Gr05Auto(bEnable := TRUE);			(* Call Program *)
Gr05Home(bEnable := TRUE);			(* Call Program *)
Gr05Manual(bEnable := TRUE);			(* Call Program *)

END_PROGRAM

// ---- POUs/Machine/Group_0500 - Transport/Gr05MachineMode/Gr05Auto/Gr05Auto.TcPOU
PROGRAM Gr05Auto
VAR_INPUT
	(* Input variables / Eingang Variablen *)
	bEnable					:BOOL;						(* Enable Gr05Auto *)
	bExecute				:BOOL;						(* Auto execute *)

	(* Instances *)
	fbInit						:FB_Gr05AutoInit;
	fbProcedure				:FB_Gr05AutoProcedure;

END_VAR
VAR
	(* Enummerations *)

	(* Variables *)
	SFCCurrentStepHis			:ARRAY[0..120] OF STRING;
	bClearHis						:BOOL;
	usnt : INT := 1;
	(* References *)

	(* Interfaces *)

	(* Instances *)
	rtExecute					:R_TRIG;
	fbAlarm					:FB_Gr05AutoAlarm;
END_VAR
VAR CONSTANT
	nFatalErrorMaxIdx				:INT := 0;						(* Maximal index of  using alarms *)
	nErrorMaxIdx					:INT := 2;						(* Maximal index of  using alarms *)
	nWarningMaxIdx				:INT := 1;						(* Maximal index of  using alarms *)
	nMessageMaxIdx				:INT := 0;						(* Maximal index of  using alarms *)
	nHintMaxIdx					:INT := 0;						(* Maximal index of  using alarms *)

	dnFatalErrorBaseIdentNo		:DINT := 52000;				(* Fatal error identification number *)
	dnErrorBaseIdentNo			:DINT := 52100;				(* Error identification number *)
	dnWarningBaseIdentNo		:DINT := 52200;				(* Warning identification number *)
	dnMessageBaseIdentNo		:DINT := 52300;				(* Message identification number *)
	dnHintBaseIdentNo			:DINT := 52400;				(* Hint identification number *)
END_VAR

IF NOT bEnable
THEN
    RETURN;
END_IF;

(* Check auto execute *)
bExecute := bgGr00ModeAutomatic
		     AND NOT fbInit.bFirstTime;

rtExecute(CLK := bExecute);

IF rtExecute.Q
THEN
	A_Init();
END_IF;

A_Procedure();
A_Functions();
A_Alarm();

ACTION A_Alarm:

(* Collect and execute input alarms *)
fbAlarm.stAlarmIn.arbError[0].bActive := fbProcedure.bErrorPipeBeginNoDetected;
fbAlarm.stAlarmIn.arbError[0].dnCode := dnErrorBaseIdentNo + 0;

fbAlarm.stAlarmIn.arbError[1].bActive := fbProcedure.bErrorPipeEndNoDetected;
fbAlarm.stAlarmIn.arbError[1].dnCode := dnErrorBaseIdentNo + 1;

fbAlarm.stAlarmIn.arbError[2].bActive := fbProcedure.bErrorCollisionDetected;
fbAlarm.stAlarmIn.arbError[2].dnCode := dnErrorBaseIdentNo + 2;

fbAlarm.stAlarmIn.arbWarning[0].bActive := fbProcedure.bWarningPipeBeginNoDetected;
fbAlarm.stAlarmIn.arbWarning[0].dnCode := dnWarningBaseIdentNo + 0;

fbAlarm(
	etMachineMode := etgGr00MachineMode,
	etMachineState := etgGr00MachineState,
	bNoEStop := bgGr00NoEmergencyStop,
	bConfirmAlarm := bgGr00ConfirmAlarm,
	dtDateTime := stgGr00DateTime.dtDateTime,
	nFatalErrorMaxIdx := nFatalErrorMaxIdx,
	nErrorMaxIdx := nErrorMaxIdx,
	nWarningMaxIdx := nWarningMaxIdx,
	nMessageMaxIdx := nMessageMaxIdx,
	nHintMaxIdx := nHintMaxIdx,
	bMoveInterrupted := bgGr05MoveInterrupted,
	bHomeCompleted := bgGr05HomeCompleted,
	stAlarmOut => stgGr05Alarm.stAuto
);
END_ACTION

ACTION A_Functions:

;
END_ACTION

ACTION A_Init:

(* Initializing variables *)
fbInit();
END_ACTION

ACTION A_Procedure:

(* Execute auto procedure *)
fbProcedure(
	bEnable := fbInit.bFirstTime,
	bExecute := bgGr05StartProcess,
	bInterrupt := FALSE(*NOT bgGr05StartProcess*),
	bReleaseNextStep := bgGr05StartProcess,
	bDone => bgGr05AutoCompleted,
	bInterrupted => bgGr05MoveInterrupted
);



(* This loup used to track the steps of this sequence *)
IF bClearHis THEN
	FOR usnt := 120 TO 1 BY  -1  DO
		SFCCurrentStepHis[usnt] := '' ;
	END_FOR
	bClearHis := FALSE;
ELSIF  fbProcedure.SFCCurrentStep <> SFCCurrentStepHis[0]  THEN
	FOR usnt := 120 TO 1 BY  -1  DO
		SFCCurrentStepHis[usnt] := SFCCurrentStepHis[usnt - 1] ;
	END_FOR
		SFCCurrentStepHis[0] := fbProcedure.SFCCurrentStep;
END_IF
END_ACTION

END_PROGRAM

// ---- POUs/Machine/Group_0500 - Transport/Gr05MachineMode/Gr05Home/Gr05Home.TcPOU
PROGRAM Gr05Home
VAR_INPUT
	(* Input variables / Eingang Variablen *)
	bEnable					:BOOL;						(* Enable Gr02Home *)
	bExecute				:BOOL;						(* Home execute *)

	(* Instances *)
	fbInit						:FB_Gr05HomeInit;
	fbProcedure				:FB_Gr05HomeProcedure;

	fbAxisClamp1				:FB_Gr05HomeAxisClamp1;
	fbAxisClamp2				:FB_Gr05HomeAxisClamp2;

END_VAR
VAR
	(* Enummerations *)

	(* Variables *)

	(* References *)

	(* Interfaces *)

	(* Instances *)
	rtExecute					:R_TRIG;

	fbAlarm					:FB_Gr05HomeAlarm;

END_VAR
VAR CONSTANT
	nFatalErrorMaxIdx				:INT := 0;						(* Maximal index of  using alarms *)
	nErrorMaxIdx					:INT := 2;						(* Maximal index of  using alarms *)
	nWarningMaxIdx				:INT := 0;						(* Maximal index of  using alarms *)
	nMessageMaxIdx				:INT := 0;						(* Maximal index of  using alarms *)
	nHintMaxIdx					:INT := 0;						(* Maximal index of  using alarms *)

	dnFatalErrorBaseIdentNo		:DINT := 53000;					(* Fatal error identification number *)
	dnErrorBaseIdentNo			:DINT := 53100;					(* Error identification number *)	
	dnWarningBaseIdentNo		:DINT := 53200;					(* Warning identification number *)	
	dnMessageBaseIdentNo		:DINT := 53300;					(* Message identification number *)	
	dnHintBaseIdentNo			:DINT := 53400;					(* Hint identification number *)
END_VAR

IF NOT bEnable
THEN
	RETURN;
END_IF;

(* Check home execute *)
bExecute := etgGr00MachineState = ET_MachineState_eHomeRefExe
		      OR etgGr00MachineState = ET_MachineState_eHomeExe;

rtExecute(CLK := bExecute);

IF rtExecute.Q
THEN
	fbInit.bFirstTime := FALSE;
	A_Init();
END_IF;

A_Procedure();
A_Functions();
A_Alarm();

ACTION A_Alarm:

(* Collect and execute input alarms *)
fbAlarm.stAlarmIn.arbError[0].bActive := fbAxisClamp1.bErrorByReference;
fbAlarm.stAlarmIn.arbError[0].dnCode := dnErrorBaseIdentNo + 0;

fbAlarm.stAlarmIn.arbError[1].bActive := fbAxisClamp1.bErrorByPipeCollision ;
fbAlarm.stAlarmIn.arbError[1].dnCode := dnErrorBaseIdentNo + 1;

fbAlarm.stAlarmIn.arbError[2].bActive := fbAxisClamp1.bErrorByPipeEndNoDetected;
fbAlarm.stAlarmIn.arbError[2].dnCode := dnErrorBaseIdentNo + 2;

fbAlarm(
	etMachineMode := etgGr00MachineMode,
	etMachineState := etgGr00MachineState,
	bNoEStop := bgGr00NoEmergencyStop,
	bConfirmAlarm := bgGr00ConfirmAlarm,
	dtDateTime := stgGr00DateTime.dtDateTime,
	nFatalErrorMaxIdx := nFatalErrorMaxIdx,
	nErrorMaxIdx := nErrorMaxIdx,
	nWarningMaxIdx := nWarningMaxIdx,
	nMessageMaxIdx := nMessageMaxIdx,
	nHintMaxIdx := nHintMaxIdx,
	bMoveInterrupted := bgGr05MoveInterrupted,
	bHomeCompleted := bgGr05HomeCompleted,
	stAlarmOut => stgGr05Alarm.stHome
);
END_ACTION

ACTION A_Functions:

fbAxisClamp1(
	bEnable := etgGr00MachineMode = ET_MachineMode_eHome,
	bReleaseNextStep := etgGr00MachineState = ET_MachineState_eHomeRefExe
		      	     		      OR etgGr00MachineState = ET_MachineState_eHomeExe
);

fbAxisClamp2(
	bEnable := etgGr00MachineMode = ET_MachineMode_eHome,
	bReleaseNextStep := etgGr00MachineState = ET_MachineState_eHomeRefExe
		      	     		      OR etgGr00MachineState = ET_MachineState_eHomeExe
);
END_ACTION

ACTION A_Init:

(* Initializing variables *)
fbInit();
END_ACTION

ACTION A_Procedure:

(* Execute home procedure *)
fbProcedure(
	bEnable := etgGr00MachineMode = ET_MachineMode_eHome,
	bExecute := rtExecute.Q,
	bReleaseNextStep := etgGr00MachineState = ET_MachineState_eHomeRefExe
		      	     		      OR etgGr00MachineState = ET_MachineState_eHomeExe
);
END_ACTION

END_PROGRAM

// ---- POUs/Machine/Group_0500 - Transport/Gr05MachineMode/Gr05Manual/Gr05Manual.TcPOU
PROGRAM Gr05Manual
VAR_INPUT
	(* Input variables / Eingang Variablen *)
	bEnable					:BOOL;						(* Enable Gr05Manual *)
	bExecute				:BOOL;						(* Manual execute *)

	(* Instances *)
	fbInit						:FB_Gr05ManualInit;
	fbProcedure				:FB_Gr05ManualProcedure;
END_VAR
VAR
	(* Enummerations *)

	(* Variables *)

	(* References *)

	(* Interfaces *)

	(* Instances *)
	rtExecute					:R_TRIG;

	fbAlarm					:FB_Gr05ManualAlarm;
END_VAR
VAR CONSTANT
	nFatalErrorMaxIdx				:INT := 0;						(* Maximal index of  using alarms *)
	nErrorMaxIdx					:INT := 0;						(* Maximal index of  using alarms *)
	nWarningMaxIdx				:INT := 0;						(* Maximal index of  using alarms *)
	nMessageMaxIdx				:INT := 0;						(* Maximal index of  using alarms *)
	nHintMaxIdx					:INT := 0;						(* Maximal index of  using alarms *)

	dnFatalErrorBaseIdentNo		:DINT := 54000;					(* Fatal error identification number *)
	dnErrorBaseIdentNo			:DINT := 54100;					(* Error identification number *)	
	dnWarningBaseIdentNo		:DINT := 54200;					(* Warning identification number *)	
	dnMessageBaseIdentNo		:DINT := 54300;					(* Message identification number *)	
	dnHintBaseIdentNo			:DINT := 54400;					(* Hint identification number *)
END_VAR

IF NOT bEnable
THEN
	RETURN;
END_IF;

(* Check manual execute *)
bExecute := etgGr00MachineMode = ET_MachineMode_eManual;

rtExecute(CLK := bExecute);

IF rtExecute.Q
THEN
	fbInit.bFirstTime := FALSE;
	A_Init();
END_IF;

A_Procedure();
A_Alarm();

ACTION A_Alarm:

(* Collect and execute input alarms *)
fbAlarm.stAlarmIn.arbError[0].bActive := FALSE;
fbAlarm.stAlarmIn.arbError[0].dnCode := dnErrorBaseIdentNo + 0;

fbAlarm(
	etMachineMode := etgGr00MachineMode,
	etMachineState := etgGr00MachineState,
	bNoEStop := bgGr00NoEmergencyStop,
	bConfirmAlarm := bgGr00ConfirmAlarm,
	dtDateTime := stgGr00DateTime.dtDateTime,
	nFatalErrorMaxIdx := nFatalErrorMaxIdx,
	nErrorMaxIdx := nErrorMaxIdx,
	nWarningMaxIdx := nWarningMaxIdx,
	nMessageMaxIdx := nMessageMaxIdx,
	nHintMaxIdx := nHintMaxIdx,
	bHomeCompleted := bgGr05HomeCompleted,
	stAlarmOut => stgGr05Alarm.stManual
);
END_ACTION

ACTION A_Init:

(* Initializing variables *)
fbInit();
END_ACTION

ACTION A_Procedure:

(* Execute manual procedure *)
fbProcedure(
	bEnable := etgGr00MachineMode = ET_MachineMode_eManual,
	bExecute := rtExecute.Q,
	bReleaseNextStep := etgGr00MachineMode = ET_MachineMode_eManual
);
END_ACTION

END_PROGRAM

// ---- POUs/Machine/Group_0500 - Transport/Gr05Control/Gr05Control.TcPOU
PROGRAM Gr05Control
VAR_INPUT
	(* Input variables / Eingang Variablen *)
	bEnable						:BOOL;						(* Enable Gr05Control *)

	(* Instances *)
	fbAxisClamp1				:FB_Gr05AxisClamp;

	arfbCylinderClamp			:ARRAY[1..ungGr05ClampMaxNo] OF FB_Gr05CylinderClamp;
	fbCylinderPos				:FB_Gr05CylinderPos;

	fbSlide						:FB_Gr05Slide;
	fbRemovalBand				:FB_Gr05RemovalBand;

END_VAR
VAR
	(* Enummerations *)

	(* Variables *)
	unClampIdx					:UINT;						(* Clamp index *)
	unCylinderPosIdx			:UINT;						(* Position cylinder index *)

	arlrAxisClampLastPos		:ARRAY[1..ungGr05ClampMaxNo] OF LREAL;

	bAllAxisCtrlEnabled			:BOOL;						(* All axis have controller enabled *)
	bAllAxisStandStill			:BOOL;						(* All axis stand still *)
	bAllAxisNotMoving			:BOOL;						(* All axis not moving *)
	bAllAxisReferenced			:BOOL;						(* All axis referenced *)

	(* References *)

	(* Interfaces *)

	(* Instances *)
	fbAlarm						:FB_Gr05Alarm;
	fbSafety					:FB_Gr05Safety;
	fbSignals					:FB_Gr05Signals;
	fbUtility					:FB_Gr05Utility;
	rtBtnStart					:R_TRIG;
	tonSlideMoveToWork			:TON;
	tpTransportBand				:TP;
END_VAR
VAR CONSTANT
	nFatalErrorMaxIdx			:INT := 0;						(* Maximal index of  using alarms *)
	nErrorMaxIdx				:INT := 23;					(* Maximal index of  using alarms *)
	nWarningMaxIdx				:INT := 0;						(* Maximal index of  using alarms *)
	nMessageMaxIdx				:INT := 3;						(* Maximal index of  using alarms *)
	nHintMaxIdx					:INT := 0;						(* Maximal index of  using alarms *)

	dnFatalErrorBaseIdentNo		:DINT := 51000;				(* Fatal error identification number *)
	dnErrorBaseIdentNo			:DINT := 51100;				(* Error identification number *)
	dnWarningBaseIdentNo		:DINT := 51200;				(* Warning identification number *)
	dnMessageBaseIdentNo		:DINT := 51300;				(* Message identification number *)
	dnHintBaseIdentNo			:DINT := 51400;				(* Hint identification number *)
END_VAR

IF NOT bEnable
THEN
	RETURN;
END_IF;

A_Utility();
A_Safety();
A_Transport();
A_Signals();
A_Alarm();

ACTION A_Alarm:

(* Collect and execute input alarms *)
fbAlarm.stAlarmIn.arbError[0].bActive := NOT binGr05LightCurtainOK
                                                		      AND (Gr05Home.fbProcedure.bBusy
                                                      				OR Gr05Auto.fbProcedure.bBusy);
fbAlarm.stAlarmIn.arbError[0].dnCode := dnErrorBaseIdentNo + 0;

fbAlarm.stAlarmIn.arbError[1].bActive := FALSE;(*(bgGr05PipeEndPresent
						       OR (bgGr05PipeBeginPresent AND Gr05Home.fbProcedure.bDone))
			                                   AND ((etgGr00MachineMode = ET_MachineMode_eHome
			                                                 AND (etgGr00MachineState = ET_MachineState_eHomeExe
			                                                      	     OR etgGr00MachineState = ET_MachineState_eHomeRefExe)))*);
fbAlarm.stAlarmIn.arbError[1].dnCode := dnErrorBaseIdentNo + 1;

fbAlarm.stAlarmIn.arbError[2].bActive := FALSE;
fbAlarm.stAlarmIn.arbError[2].dnCode := dnErrorBaseIdentNo + 2;

fbAlarm.stAlarmIn.arbError[3].bActive := FALSE;
fbAlarm.stAlarmIn.arbError[3].dnCode := dnErrorBaseIdentNo + 3;

fbAlarm.stAlarmIn.arbError[4].bActive := fbAxisClamp1.bErrorTerminal;
fbAlarm.stAlarmIn.arbError[4].dnCode := dnErrorBaseIdentNo + 4;

fbAlarm.stAlarmIn.arbError[5].bActive := fbAxisClamp1.fbController.bErrorInit;
fbAlarm.stAlarmIn.arbError[5].dnCode := dnErrorBaseIdentNo + 5;

fbAlarm.stAlarmIn.arbError[6].bActive := fbAxisClamp1.bErrorCtrlEnabled;
fbAlarm.stAlarmIn.arbError[6].dnCode := dnErrorBaseIdentNo + 6;

fbAlarm.stAlarmIn.arbError[7].bActive := fbAxisClamp1.fbController.bError OR fbAxisClamp1.fbMoveManual.bError OR fbAxisClamp1.fbMoveAuto.bError;
fbAlarm.stAlarmIn.arbError[7].dnCode := dnErrorBaseIdentNo + 7;

fbAlarm.stAlarmIn.arbError[8].bActive := arfbCylinderClamp[1].bErrorOpen;
fbAlarm.stAlarmIn.arbError[8].dnCode := dnErrorBaseIdentNo + 8;

fbAlarm.stAlarmIn.arbError[9].bActive := arfbCylinderClamp[1].bErrorClose;
fbAlarm.stAlarmIn.arbError[9].dnCode := dnErrorBaseIdentNo + 9;

fbAlarm.stAlarmIn.arbError[10].bActive := arfbCylinderClamp[2].bErrorOpen;
fbAlarm.stAlarmIn.arbError[10].dnCode := dnErrorBaseIdentNo + 10;

fbAlarm.stAlarmIn.arbError[11].bActive := arfbCylinderClamp[2].bErrorClose;
fbAlarm.stAlarmIn.arbError[11].dnCode := dnErrorBaseIdentNo + 11;

fbAlarm.stAlarmIn.arbError[12].bActive := fbSlide.bErrorMoveToBase;
fbAlarm.stAlarmIn.arbError[12].dnCode := dnErrorBaseIdentNo + 12;

fbAlarm.stAlarmIn.arbError[13].bActive := fbSlide.bErrorMoveToWork;
fbAlarm.stAlarmIn.arbError[13].dnCode := dnErrorBaseIdentNo + 13;

fbAlarm.stAlarmIn.arbError[14].bActive := fbRemovalBand.bErrorMoveToPlus;
fbAlarm.stAlarmIn.arbError[14].dnCode := dnErrorBaseIdentNo + 14;

fbAlarm.stAlarmIn.arbError[15].bActive := fbRemovalBand.bErrorMoveToMinus;
fbAlarm.stAlarmIn.arbError[15].dnCode := dnErrorBaseIdentNo + 15;

fbAlarm.stAlarmIn.arbError[16].bActive := fbRemovalBand.fbMotor.bError
						         AND fbRemovalBand.fbMotor.udnErrorNo = 8;
fbAlarm.stAlarmIn.arbError[16].dnCode := dnErrorBaseIdentNo + 16;

fbAlarm.stAlarmIn.arbError[17].bActive := fbCylinderPos.arbErrorMoveToBase[1];
fbAlarm.stAlarmIn.arbError[17].dnCode := dnErrorBaseIdentNo + 17;

fbAlarm.stAlarmIn.arbError[18].bActive := fbCylinderPos.arbErrorMoveToWork[1];
fbAlarm.stAlarmIn.arbError[18].dnCode := dnErrorBaseIdentNo + 18;

fbAlarm.stAlarmIn.arbError[19].bActive := fbCylinderPos.arbErrorMoveToBase[2];
fbAlarm.stAlarmIn.arbError[19].dnCode := dnErrorBaseIdentNo + 19;

fbAlarm.stAlarmIn.arbError[20].bActive := fbCylinderPos.arbErrorMoveToWork[2];
fbAlarm.stAlarmIn.arbError[20].dnCode := dnErrorBaseIdentNo + 20;

fbAlarm.stAlarmIn.arbError[21].bActive := fbCylinderPos.arbErrorMoveToBase[3];
fbAlarm.stAlarmIn.arbError[21].dnCode := dnErrorBaseIdentNo + 21;

fbAlarm.stAlarmIn.arbError[22].bActive := fbCylinderPos.arbErrorMoveToWork[3];
fbAlarm.stAlarmIn.arbError[22].dnCode := dnErrorBaseIdentNo + 22;

fbAlarm.stAlarmIn.arbWarning[0].bActive := FALSE;
fbAlarm.stAlarmIn.arbWarning[0].dnCode := dnWarningBaseIdentNo + 0;

fbAlarm.stAlarmIn.arbMessage[0].bActive := NOT binGr05LightCurtainOK
							      AND NOT fbAlarm.stAlarmIn.arbError[0].bActive
							      AND NOT fbAlarm.stAlarmOut.arbError[0].bActive;
fbAlarm.stAlarmIn.arbMessage[0].dnCode := dnMessageBaseIdentNo + 0;

fbAlarm.stAlarmIn.arbMessage[1].bActive := FALSE;(*bgGr05PipeEndPresent
							       AND NOT fbAlarm.stAlarmIn.arbError[1]
							       AND etgGr00MachineMode = ET_MachineMode_eHome*);
fbAlarm.stAlarmIn.arbMessage[1].dnCode := dnMessageBaseIdentNo + 1;

fbAlarm.stAlarmIn.arbMessage[2].bActive := NOT bgGr05PipeEndPresent
							      AND NOT bgGr00MachineRunning
							      AND NOT Gr05Auto.fbAlarm.stAlarmIn.arbError[0].bActive
							      AND NOT Gr05Auto.fbAlarm.stAlarmIn.arbError[1].bActive
							      AND NOT Gr05Auto.fbAlarm.stAlarmIn.arbError[2].bActive
							      AND NOT Gr05Home.fbAlarm.stAlarmOut.arbError[1].bActive
							      AND NOT Gr05Home.fbAlarm.stAlarmOut.arbError[2].bActive;
fbAlarm.stAlarmIn.arbMessage[2].dnCode := dnMessageBaseIdentNo + 2;

fbAlarm.stAlarmIn.arbMessage[3].bActive := stgGr05HMI.stPLCTOHMI.arlrAxisClampActPos[2] >= ABS(99999.0);
fbAlarm.stAlarmIn.arbMessage[3].dnCode := dnMessageBaseIdentNo + 3;


(* Execute utility *)
fbAlarm(
	etMachineMode := etgGr00MachineMode,
	etMachineState := etgGr00MachineState,
	bNoEStop := bgGr00NoEmergencyStop,
	bConfirmAlarm := bgGr00ConfirmAlarm,
	dtDateTime := stgGr00DateTime.dtDateTime,
	nFatalErrorMaxIdx := nFatalErrorMaxIdx,
	nErrorMaxIdx := nErrorMaxIdx,
	nWarningMaxIdx := nWarningMaxIdx,
	nMessageMaxIdx := nMessageMaxIdx,
	nHintMaxIdx := nHintMaxIdx,
	bMoveInterrupted := bgGr05MoveInterrupted,
	bHomeCompleted := bgGr05HomeCompleted,
	stAlarmOut => stgGr05Alarm.stControl
);
END_ACTION

ACTION A_Safety:

(* Execute safety *)
fbSafety(
	bLightCurtain := binGr05LightCurtainOK,
	bConfirmLightCurtain := (bgGr00ConfirmAlarm
			                            OR etgGr00MachineMode = ET_MachineMode_eManual
			                            OR etgGr00MachineMode = ET_MachineMode_eHome
			                            OR etgGr00MachineMode = ET_MachineMode_eAutomatic
			                            OR stgGr00HMI.stHMITOPLC.bSafetyInterlockOff)
					         AND NOT stgGr05Alarm.stControl.arbError[0].bActive,
	tLightCurtainDelay := tgGr05LightCurtainDelay,
	bLightCurtainOK => bgGr05LightCurtainOK,
	bConfirmedLightCurtain => boutGr05ConfLightCurtain
);

bgGr05SafetyActive := fbAxisClamp1.bSafetyLock;
END_ACTION

ACTION A_Signals:

(* Execute signals *)
fbSignals(
	etMachineMode := etgGr00MachineMode,
	etMachineState := etgGr00MachineState,
	bMachineRunning := bgGr00MachineRunning,
	bExecutedProcess := fbUtility.bExeProcess,
	stBlinker := stgGr00Blinker,
	bBulbBtnStart => boutGr05BulbBtnStart,
	bBulbBtnStop => boutGr05BulbBtnStop
);

(* Detect all axis controller enabled *)
bAllAxisCtrlEnabled := F_ChkAllAxisEnabled(
	bEnable := TRUE,
	bEnabledAxis1 := Gr05Control.fbAxisClamp1.bCtrlEnabled,
	bEnabledAxis2 := TRUE,
	bEnabledAxis3 := TRUE,
	bEnabledAxis4 := TRUE,
	bEnabledAxis5 := TRUE,
	bEnabledAxis6 := TRUE,
	bEnabledAxis7 := TRUE,
	bEnabledAxis8 := TRUE,
	bEnabledAxis9 := TRUE,
	bEnabledAxis10 := TRUE
);

(* Detect all axis stand still *)
bAllAxisStandStill := F_ChkAllAxisStandStill(
	bEnable := TRUE,
	bAxis1StandStill := igGr05AxisClamp1.Status.StandStill,
	bAxis2StandStill := TRUE,
	bAxis3StandStill := TRUE,
	bAxis4StandStill := TRUE,
	bAxis5StandStill := TRUE,
	bAxis6StandStill := TRUE,
	bAxis7StandStill := TRUE,
	bAxis8StandStill := TRUE,
	bAxis9StandStill := TRUE,
	bAxis10StandStill := TRUE,
);

(* Detect all axis not moving *)
bAllAxisNotMoving := F_ChkAllAxisNotMoving(
	bEnable := TRUE,
	bAxis1NotMoving := Gr05Control.fbAxisClamp1.bNotMoving, 
	bAxis2NotMoving := TRUE,
	bAxis3NotMoving := TRUE,
	bAxis4NotMoving := TRUE,
	bAxis5NotMoving := TRUE,
	bAxis6NotMoving := TRUE,
	bAxis7NotMoving := TRUE,
	bAxis8NotMoving := TRUE,
	bAxis9NotMoving := TRUE,
	bAxis10NotMoving := TRUE
);

(* Detect all axis referenced *)
bAllAxisReferenced := F_ChkAllAxisReferenced(
	bEnable := TRUE,
	bReferencedAxis1 := Gr05Control.fbAxisClamp1.bReferenced,
	bReferencedAxis2 := TRUE,
	bReferencedAxis3 := TRUE,
	bReferencedAxis4 := TRUE,
	bReferencedAxis5 := TRUE,
	bReferencedAxis6 := TRUE,
	bReferencedAxis7 := TRUE,
	bReferencedAxis8 := TRUE,
	bReferencedAxis9 := TRUE,
	bReferencedAxis10 := TRUE
);
END_ACTION

ACTION A_Transport:

(* Enable axis clamp *)
IF bgGr00ModeManual
	AND stgGr05HMI.stPLCTOHMI.arlrAxisClampActPos[2] < ABS(99999.0)
	THEN
		stgGr05HMI.stHMITOPLC.arlrAxisClampSoftLimitMin[1] := stgGr05HMI.stPLCTOHMI.arlrAxisClampActPos[2]
														+ lrgGr05CylinderPosOriginShiftPos
													   	+ lrgGr05Clamp2Width - 0.5 ;
	ELSE
		stgGr05HMI.stHMITOPLC.arlrAxisClampSoftLimitMin[1] := lrgGr05CylinderPosOriginShiftPos
												    		+ lrgGr05Clamp2Width - 0.5  ;
END_IF

lrgGr05SafetyDistance := SEL(Gr01Persistent.rPipeDiameter > 400 , 0.0 ,200.0);

stgGr05HMI.stHMITOPLC.arlrAxisClampNoRefVelo[1] := 10;

fbAxisClamp1(
	bEnable						:= TRUE,
	etMachineMode				:= etgGr00MachineMode,
	etMachineState				:= etgGr00MachineState,
	bMachineStandstill			:= bgGr00MachineStandstill,
	bNoEStop					:= bgGr00NoEmergencyStop,
	bPowerSupplyOn				:= bgGr00PowerSupplyOk,
	bSafetyOK					:= bgGr05LightCurtainOK
								   AND bgGr00AllDoorsClosedLocked,
	bCtrlInterrupt				:= FALSE,
	bMoveRelease				:= TRUE,
	bMoveInterrupt				:= FALSE,
	bPlusRelease				:= TRUE,
	bMinusRelease				:= TRUE,	(*stgGr00HMI.stHMITOPLC.bSafetyInterlockOff*)
	bSignalReference			:= NOT binGr05AxisClamp1LimitMax,
	bHWSignalLimitMax			:= NOT binGr05AxisClamp1LimitMax,
	bHWSignalLimitMin			:= NOT binGr05AxisClamp1LimitMin,
	lrSoftLimitMax				:= SEL(bgGr00ModeAutomatic, stgGr05HMI.stHMITOPLC.arlrAxisClampSoftLimitMax[1], stgGr05HMI.stHMITOPLC.arlrAxisClampSoftLimitMax[1] + 0.5),
	lrSoftLimitMin				:= SEL(bgGr00ModeAutomatic, stgGr05HMI.stHMITOPLC.arlrAxisClampSoftLimitMin[1], stgGr05HMI.stHMITOPLC.arlrAxisClampSoftLimitMin[1] - 0.5),
	bConfirmAlarm				:= bgGr00ConfirmAlarm,
	bTipPlus					:= stgGr05HMI.stHMITOPLC.arbBtnAxisClampPlus[1],
	bTipMinus					:= stgGr05HMI.stHMITOPLC.arbBtnAxisClampMinus[1],
	lrTipDistance				:= 0,
	lrManualVelocity			:= stgGr05HMI.stHMITOPLC.arlrAxisClampManualVelo[1],
	lrVelocityNoRef				:= stgGr05HMI.stHMITOPLC.arlrAxisClampNoRefVelo[1],
	bVelocityLimitEn			:= FALSE,
	lrAcceleration				:= 100.0,
	lrDeceleration				:= 100.0,
	lrJerk						:= 100.0,
	lrOverride					:= fbUtility.rActOverride,
	lrExtOverride				:= 100.0,
	dnRatioNumerator			:= 1,
	udnRatioDenominator			:= 1,
	bEngineTorqueLimitEn		:= FALSE,
	lrEngineTorque				:= 200.0,
	tControllerOff				:= tgGr05ControllerOff,
	bWithAbsoluteEncoder		:= FALSE,
	lrOriginShift				:= stgGr05HMI.stHMITOPLC.arlrAxisClampOriginShiftPos[1],
	bVeloForceCtrlEn			:= FALSE,
	tAdsTimeOut					:= DEFAULT_ADS_TIMEOUT,
	bHomeCompleted				:= bgGr05HomeCompleted,
	Drive						:= igGr05DriveClamp1,
	Axis						:= igGr05AxisClamp1,
	MasterAxis					:= GVL_Gr00Interface.iAxisDummy,
	lrActPosition				=> stgGr05HMI.stPLCTOHMI.arlrAxisClampActPos[1],
	lrActVelocity				=> stgGr05HMI.stPLCTOHMI.arlrAxisClampActVelo[1],
	lrActForce					=> stgGr05HMI.stPLCTOHMI.arlrAxisClampActForce[1]
);


(* Control open/close clamp cylinder *)
FOR unClampIdx :=1 TO ungGr05ClampMaxNo
DO
	arfbCylinderClamp[unClampIdx](
		etMachineMode := etgGr00MachineMode,
		etMachineState := etgGr00MachineState,
		bAirPressureOK := bgGr00AirPressureOK,
		bSafetyOK := bgGr05LightCurtainOK
				        AND bgGr00AllDoorsClosedLocked,
		bOpened := arbinGr05ClampOpened[unClampIdx],
		bClosed := arbinGr05ClampClosed[unClampIdx],
		bHandOpen := stgGr05HMI.stHMITOPLC.arbBtnClampOpen[unClampIdx],
		bHandClose := stgGr05HMI.stHMITOPLC.arbBtnClampClose[unClampIdx],
		bOpenRelease := TRUE,
		bCloseRelease := TRUE,
		bControlOff := NOT bgGr00NoEmergencyStop,
		bConfirmAlarm := bgGr00ConfirmAlarm,
		tTimeOut := t#15s,
		bHomeCompleted := bgGr05HomeCompleted,
		bOpen => arboutGr05ClampOpen[unClampIdx],
		bClose => arboutGr05ClampClose[unClampIdx]
	);

END_FOR

(* Control position cylinder *)
stgGr05HMI.stHMITOPLC.bCylinderPosActive := TRUE;

fbCylinderPos(
	bEnable := stgGr05HMI.stHMITOPLC.bCylinderPosActive,
	etMachineMode := etgGr00MachineMode,
	etMachineState := etgGr00MachineState,
	bNoEStop := bgGr00NoEmergencyStop,
	bSafetyOK := bgGr05LightCurtainOK
			        AND bgGr00AllDoorsClosedLocked,
	bAirPressureOK := bgGr00AirPressureOK,
	lrPosOffset := lrgGr05CylinderPosOffset,
	lrOriginShiftPos := lrgGr05CylinderPosOriginShiftPos,
	etDirection := etgGr05CylinderPosDirection,
	usnCodingType := usngGr05CylinderPosCodingType,
	bControlOff := FALSE,
	bConfirmAlarm := bgGr00ConfirmAlarm,
	tTimeOut := t#10s,
	bHomeCompleted := bgGr05HomeCompleted,
	lrActPosition => stgGr05HMI.stPLCTOHMI.arlrAxisClampActPos[2]
 );

IF NOT stgGr05HMI.stHMITOPLC.bCylinderPosActive
     AND arlrAxisClampLastPos[2] <> stgGr05HMI.stPLCTOHMI.arlrAxisClampActPos[2]
THEN
	bgGr05HomeCompleted := FALSE;
	arlrAxisClampLastPos[2] := stgGr05HMI.stPLCTOHMI.arlrAxisClampActPos[2];
END_IF

FOR unCylinderPosIdx := 1 TO ungGr05CylinderPosMaxNo
DO
	fbCylinderPos.arbHandMoveToBase[unCylinderPosIdx] := stgGr05HMI.stHMITOPLC.arbBtnCylinderPosClose[unCylinderPosIdx];
	fbCylinderPos.arbHandMoveToWork[unCylinderPosIdx] := stgGr05HMI.stHMITOPLC.arbBtnCylinderPosOpen[unCylinderPosIdx];
	fbCylinderPos.arbInBase[unCylinderPosIdx] := arbinGr05CylinderPosClosed[unCylinderPosIdx];
	fbCylinderPos.arbInWork[unCylinderPosIdx] := arbinGr05CylinderPosOpened[unCylinderPosIdx];
	fbCylinderPos.arbMoveToBaseRelease[unCylinderPosIdx] := TRUE;
	fbCylinderPos.arbMoveToWorkRelease[unCylinderPosIdx] := TRUE;
	arboutGr05CylinderPosOpen[unCylinderPosIdx] := fbCylinderPos.arbMoveToWork[unCylinderPosIdx];
	arboutGr05CylinderPosClose[unCylinderPosIdx] := fbCylinderPos.arbMoveToBase[unCylinderPosIdx];
END_FOR

(* Control slide cylinder *)
tonSlideMoveToWork(
	IN := fbSlide.bAutoMoveToWork
		AND fbSlide.fbCylinder.bEndWork,
	PT := tgGr05SlideWaitInWork
);

IF bgGr00ModeAutomatic
     AND bgGr00MachineRunning
     AND tonSlideMoveToWork.Q
THEN
	fbSlide.bAutoMoveToBase := TRUE;
	fbSlide.bAutoMoveToWork := FALSE;
END_IF

stgGr05HMI.stHMITOPLC.bSlideActive := FALSE;

fbSlide(
	bEnable := stgGr05HMI.stHMITOPLC.bSlideActive,
	etMachineMode := etgGr00MachineMode,
	etMachineState := etgGr00MachineState,
	bAirPressureOK := bgGr00AirPressureOK,
	bSafetyOK := bgGr05LightCurtainOK
			        AND bgGr00AllDoorsClosedLocked,
	bInBase := binGr05SlideTop,
	bInWork := binGr05SlideBottom,
	bMoveToBaseRelease := TRUE,
	bMoveToWorkRelease := TRUE,
	bHandMoveToBase := stgGr05HMI.stHMITOPLC.bBtnSlideUp,
	bHandMoveToWork := stgGr05HMI.stHMITOPLC.bBtnSlideDown,
	bControlOff := NOT bgGr00NoEmergencyStop,
	bConfirmAlarm := bgGr00ConfirmAlarm,
	tTimeOut := t#6s,
	bHomeCompleted := bgGr05HomeCompleted,
	bMoveToBase => boutGr05SlideUp,
	bMoveToWork => boutGr05SlideDown
);

(* Control removal band *)
tpTransportBand(IN := Gr05Home.bExecute, PT := t#5s);

fbRemovalBand.arbAutoMoveToMinus[1] := binGr05PushBtnRemovalBandStart
									    OR tpTransportBand.Q
									    OR (fbAxisClamp1.lrActVelocity < 0.0 AND NOT fbAxisClamp1.bNotMoving);

IF NOT bgGr00MachineRunning
THEN
	fbRemovalBand.arbAutoMoveToMinus[2] := FALSE;
END_IF

fbRemovalBand(
	etMachineMode := etgGr00MachineMode,
	etMachineMode := etgGr00MachineMode,
	etMachineState := etgGr00MachineState,
	bNoEStop := bgGr00NoEmergencyStop,
	bPowerSupplyOn := bgGr00PowerSupplyOk
					   AND NOT binGr05RemovalBandNOK,
	bSafetyOK := bgGr05LightCurtainOK
			        AND bgGr00AllDoorsClosedLocked,
	bInPlusLimit := binGr05RemovalBandInPlus,
	bInMinusLimit := binGr05RemovalBandInMinus,
	bMoveToPlusRelease := NOT binGr05RemovalBandNOK,
	bMoveToMinusRelease := NOT binGr05RemovalBandNOK,
	bHandMoveToPlus := stgGr05HMI.stHMITOPLC.bBtnRemovalBandToPlus,
	bHandMoveToMinus := binGr05PushBtnRemovalBandStart
					        OR stgGr05HMI.stHMITOPLC.bBtnRemovalBandToMinus
					        OR (fbAxisClamp1.lrActVelocity < 0.0 AND NOT fbAxisClamp1.bNotMoving),
	bAutoMoveToPlus := FALSE,
	bConfirmAlarm := bgGr00ConfirmAlarm,
	tTimeOut := t#6s,
	bHomeCompleted := bgGr05HomeCompleted,
	bMoveToPlus => boutGr05RemovalBandToPlus,
	bMoveToMinus => boutGr05RemovalBandToMinus
);
END_ACTION

ACTION A_Utility:

(* Execute utility *)
rtBtnStart(CLK := binGr00PushBtnStart OR stgGr00HMI.stHMITOPLC.bBtnStart);

fbUtility(
	etMachineMode := etgGr00MachineMode,
	etMachineState := etgGr00MachineState,
	bStartProcess := (*stgGr05HMI.stHMITOPLC.bBtnStart*)
					rtBtnStart.Q
					AND etgGr00MachineState = ET_MachineState_eAutoExe,
	bStopProcess := (*stgGr05HMI.stHMITOPLC.bBtnStop*)
				       etgGr00MachineState <> ET_MachineState_eAutoExe,
	bSteppingProcess := stgGr05HMI.stHMITOPLC.bBtnSteppingProcess,
	bAutoCompleted := bgGr00AutoCompleted
					  AND bgGr01AutoCompleted
					  AND bgGr05AutoCompleted
					  AND bgGr05AutoCompleted
					  AND bgGr00MachineStandstill
					  AND etgGr00MachineState <> ET_MachineState_eAutoExe,
	bHomeCompleted := bgGr05HomeCompleted,
	bExeCounter := bgGr05AutoCompleted,
	bStartTime :=  fbUtility.bStartProcess,
	bStopTime := bgGr05AutoCompleted
				OR fbUtility.bStopProcess,
	bLifetimeOn := FALSE,
	bResetLifetimeAll := FALSE,
	bResetLifetime := stgGr05HMI.stHMITOPLC.bResetLifetime,
	sLifetimeFilePath := sgGr05LifetimeFilePath,
	sLifetimeFileName := sgGr05LifetimeFileName,
	bPipeEndEdgeIdentify := binGr05PipeEndEdge,
	bPipeBeginEdgeIdentify := binGr05PipeBeginEdge,
	rGlobalOverride := rgGr00Override,
	rLocalOverride := stgGr05HMI.stHMITOPLC.rOverride,
	lrLifetimeAll => stgGr05HMI.stPLCTOHMI.lrLifetime,
	lrLifetimeAfterReset => stgGr05HMI.stPLCTOHMI.lrLifetimeAfterReset,
	lrLifetimeAfterTrunOn => stgGr05HMI.stPLCTOHMI.lrLifetimeAfterTurnOn,
	udnCounterTotal := stgGr05HMI.stPLCTOHMI.udnCounterTotal,
	tAdsTimeOut := DEFAULT_ADS_TIMEOUT,
	bExeProcess => bgGr05StartProcess,
	bPipeEndPresent => bgGr05PipeEndPresent,
	bPipeBeginPresent => bgGr05PipeBeginPresent
);
END_ACTION

END_PROGRAM

// ---- POUs/Machine/Group_0500 - Transport/Gr05Control/Gr05Units/FB_Gr05AxisClamp.TcPOU
FUNCTION_BLOCK FB_Gr05AxisClamp
(*

The function block used to control axis Clamp.

Constructor: 		Patryk Panylo
Company:		E. Riexinger GmbH
Date:			28.04.2015
Version:			1.00

Date:			Revision:		Who:				Comment
dd.mm.yyyy		x.xx			Initials			comment

*)
VAR_INPUT
	(* Input variables / Eingang Variablen *)

	(* --- Axis / Achse --- *)
	bEnable						:BOOL;						(* Axis present *)

	(* --- Machine state / Maschinenzustand --- *)
	etMachineMode				:ET_MachineMode;			(* Machine mode *)
	etMachineState				:ET_MachineState;			(* Machine state *)
	bMachineStandstill			:BOOL;						(* Machine standstill *)

	(* --- Safety & releases / Sicherheit & Freigaben --- *)
	bNoEStop					:BOOL;						(* No ermergency Stop / Keine Notaus *)
	bPowerSupplyOn				:BOOL;						(* Power supply on / Leitung eingeschaltet *)
	bSafetyOK					:BOOL;						(* Safety ok / Sicherheit i.o *)
	bCtrlInterrupt				:BOOL;						(* Control interrupt *)
	bMoveRelease				:BOOL;						(* Move release *)
	bMoveInterrupt				:BOOL;						(* Move Interrupt *)
	bPlusRelease				:BOOL;						(* Plus move release *)
	bMinusRelease				:BOOL;						(* Minus move release *)

	(* --- Limits & signals / Endlagen & Signale --- *)
	bSignalReference			:BOOL;						(* Reference signal *)
	bHWSignalLimitMax			:BOOL;						(* Signal position limit switch maximum *)
	bHWSignalLimitMin			:BOOL;						(* Signal position limit switch minimum *)
	lrSoftLimitMax				:LREAL;						(* Position limit switch maximum *)
	lrSoftLimitMin				:LREAL;						(* Position limit switch minimum *)

	(* --- Commands / Befehle --- *)
	bExeReset					:BOOL;						(* Execute auto reset *)
	bExeSetPos					:BOOL;						(* Execute set position *)
	bExeHome					:BOOL;						(* Execute home *)
	bExeMoveAbs					:BOOL;						(* Execute move absolut *)
	bExeMoveRel					:BOOL;						(* Execute move relative *)
	bExeMoveAdd					:BOOL;						(* Execute move additive *)
	bExeMoveSuper				:BOOL;						(* Execute move superimposed *)
	bExeMoveVelo				:BOOL;						(* Execute move velo *)
	bExeGearIn					:BOOL;						(* Execute gear in *)
	bExeGearOut					:BOOL;						(* Execute gear out *)
	bExeStop					:BOOL;						(* Execute move stop *)
	bConfirmAlarm				:BOOL;						(* Confirm alarm *)

	(* --- Manual mode / Handbetrieb --- *)
	bTipPlus					:BOOL;						(* Manual tip in plus direction *)
	bTipMinus					:BOOL;						(* Manual tip in minus direction *)
	lrTipDistance				:LREAL;						(* Relative distance for movements *)
	lrManualVelocity			:LREAL;						(* Value of velocity in manual motion [mm/s] *)

	(* --- Motion parameters / Bewegungsparameter --- *)
	lrTargetPosition			:LREAL;						(* Absolute target position *)
	lrAutoVelocity				:LREAL;						(* Value of velocity in auto motion [mm/s] *)
	lrVelocityNoRef				:LREAL;						(* Velocity if has no reference [mm/s] *)
	bVelocityLimitEn			:BOOL;						(* Enable velocity limit *)
	lrVelocityMin				:LREAL;						(* Velocity minimum [%] *)
	lrVelocityMax				:LREAL;						(* Velocity maximum [%] *)
	lrAcceleration				:LREAL;						(* Value of the acceleration (always positive) *)
	lrDeceleration				:LREAL;						(* Value of deceleration (always positive) *)
	lrJerk						:LREAL;						(* Value of jerk (always positive) *)

	(* --- Override --- *)
	lrOverride					:LREAL;						(* Override *)
	bExtOverrideEn				:BOOL;						(* External override enable *)
	lrExtOverride				:LREAL;						(* External override *)

	(* --- Gearing / Getriebe --- *)
	dnRatioNumerator			:DINT;						(* Gear ratio numerator. Alternatively, the gear ratio can be specified in the numerator as a floating comma value, if the denominator is 1. *)
	udnRatioDenominator			:UDINT;						(* Gear ratio denominator *)

	(* --- Drive / Antrieb --- *)
	snModesOfOperation			:SINT;						(* Modes of drive operation *)
	bEngineTorqueLimitEn		:BOOL;						(* Enable engine torque limit *)
	lrEngineTorque				:LREAL;						(* Engine torque [%] *)
	tControllerOff				:TIME := T#60S;				(* Time to switch controller off *)

	(* --- Encoder / Geber --- *)
	bWithAbsoluteEncoder		:BOOL;						(* Encoder is an absolute one / Absolutwertgeber *)
	lrOriginShift				:LREAL;						(* Origin shift position *)

	(* --- Force control / Kraftregelung --- *)
	unForceMeasureType			:UINT;						(* Type of force measure system. 1: Simple mA,  2: EL3351 3: EL3356 *)
	bVeloForceCtrlEn			:BOOL;						(* Enable velocity - force controller *)
	lrVeloForceCtrlKp			:LREAL;						(* Velocity - force controller proportional band Kp *)
	lrVeloForceCtrlTi			:LREAL;						(* Velocity - force controller integral Ti *)
	lrVeloForcePreCtrlVelo		:LREAL;						(* Feedforward velocity precontrol wieghting =  0..1 *)
	lrVeloForceCtrlLimit		:LREAL;						(* Velocity - force controller limit  *)
	lrTargetForce				:LREAL;						(* Absolute target force [N] *)
	lrForceCurrent				:LREAL;						(* Current force [mA] *)
	lrForceOffset				:LREAL;						(* Force offset [N] *)
	lrForceMin					:LREAL;						(* Force min 16#0000 *)
	lrForceMax					:LREAL;						(* Force max 16#7FFF *)
	lrForceMinN					:LREAL;						(* Force min [N] *)
	lrForceMaxN					:LREAL;						(* Force max [N] *)

	(* --- System --- *)
	tAdsTimeOut					:TIME := T#2S;				(* Timout for ads commands *)
END_VAR
VAR_OUTPUT
	(* Output variables / Ausgang Variablen *)

	(* --- Status --- *)
	bCtrlEnabled				:BOOL;						(* Controller enabled *)
	bNotMoving					:BOOL;						(* Axis not moving *)
	bReferenced					:BOOL;						(* Axis referenced *)
	bCoupled					:BOOL;						(* Axis coupled *)

	(* --- Actual values / Istwerte --- *)
	lrActPosition				:LREAL;						(* Actual position [mm] *)
	lrActVelocity				:LREAL;						(* Actual velocity [mm/s] *)
	lrActForce					:LREAL;						(* Actual force [N] *)

	(* --- Limits / Endlagen --- *)
	bHardLimitMaxExceeded		:BOOL;						(* Position limit switch maximum is exceeded *)
	bHardLimitMinExceeded		:BOOL;						(* Position limit switch minimum is exceeded *)
	bSoftLimitMaxExceeded		:BOOL;						(* Position limit switch maximum is exceeded *)
	bSoftLimitMinExceeded		:BOOL;						(* Position limit switch minimum is exceeded *)

	(* --- Safety / Sicherheit --- *)
	bSafetyLock					:BOOL;						(* Safety lock*)

	(* --- Errors / Fehler --- *)
	bErrorTerminal				:BOOL;						(* Error Axis terminal *)
	bErrorCtrlEnabled			:BOOL;						(* Error Axis controller enabled *)
END_VAR
VAR_IN_OUT
	(* Input Output variables / Ausgang Variablen *)
	bHomeCompleted				:BOOL;						(* Home completed *)
	Drive						:ST_STOEBERSI6SC6CIA402_REF; (* Interface NC -> PLC *)
	Axis						:AXIS_REF;					(* Interface PLC -> NC *)
	MasterAxis					:AXIS_REF;					(* Interface with Master Axis -> is no so dummy *)
END_VAR
VAR
	(* Enummerations *)

	(* Variables *)
	sAdsAddr					:STRING(23);				(* AmsNetId of the EtherCAT master device.*)
	unSlaveAddr					:UINT;						(* Address of the slave device.*)
	
	nTorqueLimitMax				:INT := 100;
	nVelocityLimitMax			:INT := 100;

	lrVeloLimitMax				:LREAL;
	lrVeloLimitMin				:LREAL;

	sTerminalStatus				:STRING;

	bSetCoeParaToDefault		:BOOL;
	bReadCoePara				:BOOL;
	bWriteCoePara				:BOOL;
	stCoeWrite					:ST_EL3356CoeInfo;
	stCoeRead					:ST_EL3356CoeInfo;

	lrCacheWeightTara			:LREAL;

	(* References *)

	(* Interfaces *)

	(* Instances *)
	fbTerminalDiagnosis			:FB_TerminalDiagnosis;
	rtMachineStandstill			:R_TRIG;
	tonAxisEnabled				:TON;

	fbController				:FB_STOEBER_AxisController;
	fbMoveManual				:FB_STOEBER_AxisMoveManual;
	fbMoveAuto					:FB_STOEBER_AxisMoveAuto;
	// fbLink						:FB_STOEBER_DriveLink;	// Was active, aber gibts doch gar nicht mehr 
	fbForceSimple				:FB_ScalingOffset;
	fbForceEL3351				:FB_EL3351;
	fbForceEL3356				:FB_EL3356;
	fbForceCtrl					:FB_ForceController;
	fbSawingOverride			:FB_Override;

	rtWriteForcePara			:R_TRIG;

END_VAR


IF NOT bEnable								(* Signal FB enable *)
THEN

	RETURN;
END_IF


A_AxisLink();
A_AxisGetStatus();
A_AxisController();
A_AxisForceCtrl();
A_AxisMoveManual();
A_AxisMoveAuto();
A_AxisTerminalDiag();
A_AxisAlarm();

ACTION A_AxisAlarm:

(* Axis error *)
tonAxisEnabled(
	IN := fbController.bEnable
		AND fbController.bRegulatorOn
		AND NOT fbController.bStatusDelay,
	PT := fbController.tStatusDelay + t#2s
);

bErrorCtrlEnabled := tonAxisEnabled.Q;
(*byErrorPLCOpenController := fbAxisControl.byPLCOpenErrCode;*)
(*bErrorController := fbAxisControl.bError;
bErrorMoveManual := fbMoveManual.bError;
bErrorMoveAuto := fbMoveAuto.bError;*)
END_ACTION

ACTION A_AxisController:

(* Axis controller *)
fbController(
    bEnable 				:= TRUE,
	etMachineMode 			:= etMachineMode,
	etMachineState 			:= etMachineState,
	bRegulatorOn 			:= 	bNoEStop
				      			AND bPowerSupplyOn
				      			AND bSafetyOK
                   		      	AND NOT bCtrlInterrupt
				     	 		AND NOT fbMoveManual.bControllerOff
				      			AND NOT fbMoveAuto.bControllerOff,
	bReset 					:= bConfirmAlarm,
	bCMDInterrupt 			:= bMoveInterrupt,
	bTerminalOK 			:= fbTerminalDiagnosis.bTerminalOK,
	bExeReset 				:= bExeReset,
  	bExeGearIn 				:= bExeGearIn,
    bExeGearOut 			:= bExeGearOut,
   	dnRatioNumerator 		:= dnRatioNumerator,
   	udnRatioDenominator 	:= udnRatioDenominator,
	lrOverride 				:= SEL(bExtOverrideEn,
									SEL(bVeloForceCtrlEn,
										lrOverride,
										fbForceCtrl.lrCVVelo),
									lrExtOverride),
	bWithAbsoluteEncoder 	:= bWithAbsoluteEncoder,
	bSignalHWLimitMax 		:= bHWSignalLimitMax,
	bSignalHWLimitMin 		:= bHWSignalLimitMin,
	lrSoftLimitMax 			:= lrSoftLimitMax,
	lrSoftLimitMin 			:= lrSoftLimitMin,
	lrAcceleration 			:= lrAcceleration,
	lrDeceleration 			:= lrDeceleration,
	lrJerk 					:= lrJerk,
	tAdsTimeOut 			:= tAdsTimeOut,
	Axis 					:= Axis,
	MasterAxis				:= MasterAxis,
	
	bStatusDelay 			=> bCtrlEnabled,
	lrActPos 				=> lrActPosition,
	lrActVelo 				=> lrActVelocity,
	bNotMoving 				=> bNotMoving,
	bReferenced 			=> bReferenced,
	bCoupled 				=> bCoupled,
	bHardLimitMaxExceeded 	=> bHardLimitMaxExceeded,
	bHardLimitMinExceeded 	=> bHardLimitMinExceeded,
	bSoftLimitMaxExceeded 	=> bSoftLimitMaxExceeded,
	bSoftLimitMinExceeded 	=> bSoftLimitMinExceeded
);
END_ACTION

ACTION A_AxisForceCtrl:

IF unForceMeasureType = 1			(* Current or voltage force measure *)
THEN
	fbForceCtrl.lrMaxForce := lrForceMaxN; (* [N] *)

	fbForceSimple(
		bEnable := TRUE,
		lrInput := lrForceCurrent,
		lrXLowLimit := lrForceMin, (* 16#0000 = 4 [mA] *)
		lrXUpperLimit := lrForceMax, (* 16#7FFF = 20 [mA] *)
		lrYLowLimit := lrForceMinN,  (*[N]*)
		lrYUpperLimit := lrForceMaxN,  (*[N]*)
		usiPrecision := 2,
		lrOffset := LREAL_TO_REAL(lrForceOffset),
		lrOutputPV => lrActForce
	);


ELSIF unForceMeasureType = 2			(* EL3351 force measure *)
THEN
	fbForceCtrl.lrMaxForce := lrForceMaxN; (* [N] *)

	fbForceEL3351(
		bEnable := TRUE,
		nTerminalNr := 1,
		stTerminalState := ,
		stBridgeState := ,
		stSupplyState := ,
		dnRefvoltage := ,
		dnDiffvoltage := ,
		rOffset := LREAL_TO_REAL(lrForceOffset),
		usiPrecision := 2,
		bDeviceOk => ,
		sDeviceStatus => ,
		rUdiff => ,
		rUref => ,
		lrGrossWeightRV=> ,
		lrGrossWeightPV => lrActForce,
		lrNetWeightRV=> ,
		lrNetWeightPV=> ,
		lrTareWeightRV=> ,
		lrTareWeightPV=>
	);

ELSIF  unForceMeasureType = 3			(* EL3356 force measure *)
THEN

(*
	rtWriteForcePara(
		CLK:= bgGr01ForceActiv5kN
			   XOR bgGr01ForceActiv10kN
	);

	CASE nStepWriteForcePara OF
		0:	(*Idle*)

			fbForceEL3356.bWriteCoePara:= FALSE;
			bWriteForceParaBusy := FALSE;

			IF rtWriteForcePara.Q
			THEN
				nStepWriteForcePara := 10;
				bWriteForceParaBusy := TRUE;
			END_IF
		10: 	(*Start*)

			IF bgGr01ForceActiv5kN
			THEN
				fbForceCtrl.lrMaxForce := 5000, (* [N] *)

				stCoeWrite.bEnableFilter := TRUE;
				stCoeWrite.bEnableUserScale := TRUE;
				stCoeWrite.dwFilterSettings := 0;
				stCoeWrite.rGain := 1.0;
				stCoeWrite.rTara := stgGr01HMI.stHMITOPLC.lrOriginShiftForceX2Right;
				stCoeWrite.rRatedOutput := 0.995000;
				stCoeWrite.rNominalLoad := 5000.0;
				stCoeWrite.rZeroBalance := -0.00028;
				stCoeWrite.rGravityOfEarth := 9.806650;
				stCoeWrite.rScaleFactor := 1.0;
				stCoeWrite.rReferenceLoad	:= 5.0;
				stCoeWrite.bEnableUserScaleIndex8010 := FALSE;
				stCoeWrite.dnUserScaleOffsetIndex8010 := 0;
				stCoeWrite.dnUserScaleGainIndex8010 := 65536;
				stCoeWrite.dwFilterSettingsIndex8010	:= 0;

				fbForceEL3356.bWriteCoePara:= TRUE;

				nStepWriteForcePara := 20;

			ELSIF bgGr01ForceActiv10kN
			THEN
				fbForceCtrl.lrMaxForce := 10000, (* [N] *)

				stCoeWrite.bEnableFilter := TRUE;
				stCoeWrite.bEnableUserScale := TRUE;
				stCoeWrite.dwFilterSettings := 0;
				stCoeWrite.rGain := 1.0;
				stCoeWrite.rTara := stgGr01HMI.stHMITOPLC.lrOriginShiftForceX2Right;
				stCoeWrite.rRatedOutput := 0.9907;
				stCoeWrite.rNominalLoad := 10000.0;
				stCoeWrite.rZeroBalance := 0.00147;
				stCoeWrite.rGravityOfEarth := 9.806650;
				stCoeWrite.rScaleFactor := 1.0;
				stCoeWrite.rReferenceLoad	:= 10.0;
				stCoeWrite.bEnableUserScaleIndex8010 := FALSE;
				stCoeWrite.dnUserScaleOffsetIndex8010 := 0;
				stCoeWrite.dnUserScaleGainIndex8010 := 65536;
				stCoeWrite.dwFilterSettingsIndex8010	:= 0;

				fbForceEL3356.bWriteCoePara:= TRUE;

				nStepWriteForcePara := 20;

			ELSE

				nStepWriteForcePara := 40;
			END_IF

		20: 	(*Wait*)
			IF fbForceEL3356.fbCoe.bCoeBusy
			THEN
				fbForceEL3356.bWriteCoePara:= FALSE;

				nStepWriteForcePara := 30;
			END_IF
	
		30: (*Write*)
			IF NOT fbForceEL3356.fbCoe.bCoeBusy
			THEN
				bWriteForceParaBusy := FALSE;

				IF NOT fbForceEL3356.fbCoe.bCoeError
				THEN
					nStepWriteForcePara := 0;
				ELSE
					nStepWriteForcePara := 40;
				END_IF
			END_IF
		40: (*Error*)
			nStepWriteForcePara := 0;

		ELSE
			nStepWriteForcePara := 0;
	END_CASE

*)

	fbForceCtrl.lrMaxForce := 5000; (* [N] *)

	stCoeWrite.bEnableFilter := TRUE;
	stCoeWrite.bEnableUserScale := TRUE;
	stCoeWrite.dwFilterSettings := 0;
	stCoeWrite.rGain := 1.0;
	stCoeWrite.rTara := (*stgGr01HMI.stHMITOPLC.lrOriginShiftForce*)0.0;
	stCoeWrite.rRatedOutput := 0.995000;
	stCoeWrite.rNominalLoad := 5000.0;
	stCoeWrite.rZeroBalance := -0.00028;
	stCoeWrite.rGravityOfEarth := 9.806650;
	stCoeWrite.rScaleFactor := 1.0;
	stCoeWrite.rReferenceLoad	:= 5.0;
	stCoeWrite.bEnableUserScaleIndex8010 := FALSE;
	stCoeWrite.dnUserScaleOffsetIndex8010 := 0;
	stCoeWrite.dnUserScaleGainIndex8010 := 65536;
	stCoeWrite.dwFilterSettingsIndex8010	:= 0;

	bWriteCoePara := lrCacheWeightTara <> (*stgGr01HMI.stHMITOPLC.lrOriginShiftForce*)0.0;

	fbForceEL3356(
		bEnable := TRUE,
		nTerminalNr := 1,
(*		stTerminalState := stinGr01EL3356A12TerminalState,
		stChannelState := stinGr01EL3356A12ChannelState,*)
		bSetCoeParaToDefault := bSetCoeParaToDefault,
		bReadCoePara := bReadCoePara,
		bWriteCoePara := bWriteCoePara,
		rValue := (*rinGr01ForceRMBValue*)0.0,
		stCoeWrite := stCoeWrite,
		stCoeRead => stCoeRead,
(*		stChannelCtrl => stoutGr01EL3356A8ChannelCtrl,*)
		lrGrossWeightPV =>
	);

	lrActForce := F_LRealRound(fbForceEL3356.lrGrossWeightPV - lrForceOffset, 2);

	lrCacheWeightTara := (*stgGr01HMI.stHMITOPLC.lrOriginShiftForce*)0.0;

ELSE							(* Directly force measure *)

	lrActForce := lrForceCurrent;
	fbForceCtrl.lrMaxForce := lrForceMaxN; (* [N] *)

END_IF

fbForceCtrl(
	bEnable := bNoEStop
			    AND bPowerSupplyOn
			    AND bSafetyOK
			    AND bCtrlEnabled,
	bControllerOn := bVeloForceCtrlEn,
	lrVeloKp := lrVeloForceCtrlKp,
	lrVeloTi := lrVeloForceCtrlTi,
	lrCtrlVeloFilter := lrVeloForcePreCtrlVelo,
	lrPVForce := lrActForce, (* [N] *)
	lrSPForce := lrTargetForce, (* [N] *)
	lrVeloMax := lrVeloForceCtrlLimit,
	lrVeloMin := -lrVeloForceCtrlLimit,
	lrTaskCycle := lrgActCycleTime
);
END_ACTION

ACTION A_AxisGetStatus:

(* Get axis status *)
Axis.ReadStatus();
END_ACTION

ACTION A_AxisLink:

(* Get terminal status *)
sAdsAddr := F_CreateAmsNetId(Drive.stTerminalState.stAdsAddr.netId);
unSlaveAddr := Drive.stTerminalState.stAdsAddr.port;
Axis.DriveAddress.NetID := F_CreateAmsNetId(Drive.stTerminalState.stAdsAddr.netId);
Axis.DriveAddress.SlaveAddress := Drive.stTerminalState.stAdsAddr.port;

(* Set drive parameter *)
Drive.stPlcToStoeber.snA541ModesOfOperation := snModesOfOperation;

(*Drive.PlcToStoeber.nA558TargetTorque := SEL(bEngineTorqueLimitEn,
				    nTorqueLimitMax,
				    LREAL_TO_INT(lrEngineTorque / 1.0))*)








(*



(* Axis linking *)
fbLink(
	Drive := Drive,
	Axis := Axis
);


*)
END_ACTION

ACTION A_AxisMoveAuto:

(* Move axis auto *)
rtMachineStandstill(CLK := bMachineStandstill);

lrVeloLimitMin := SEL(bVelocityLimitEn, INT_TO_LREAL( -1 * nVelocityLimitMax), lrVelocityMin);
lrVeloLimitMax := SEL(bVelocityLimitEn, INT_TO_LREAL(nVelocityLimitMax), lrVelocityMax);

fbMoveAuto(
	bEnable 			:= bNoEStop
               		    	AND bPowerSupplyOn
               		    	AND bSafetyOK,
    bCtrlEnabled 		:= bCtrlEnabled
                    		   AND bMoveRelease,
	etMachineMode 		:= etMachineMode,
	etMachineState 		:= etMachineState,
	bReset 				:= bConfirmAlarm,
	bExeHome 			:= bExeHome,
	bExeMoveAbs 		:= bExeMoveAbs,
	bExeMoveRel 		:= bExeMoveRel,
	bExeMoveAdd 		:= bExeMoveAdd,
	bExeMoveSuper 		:= bExeMoveSuper,
	bExeMoveVelo 		:= bExeMoveVelo,
	bExeStop 			:= bExeStop
			      			OR rtMachineStandstill.Q,
	lrPosition 			:= lrTargetPosition,
	lrVelocity 			:= LIMIT(lrVeloLimitMin, lrAutoVelocity, lrVeloLimitMax),
	lrAcceleration 		:= lrAcceleration,
	lrDeceleration 		:= lrDeceleration,
	lrJerk 				:= lrJerk,
	lrOriginShiftPos 	:= lrOriginShift,
	bSignalReference 	:= bSignalReference,
	tControllerOff 		:= tControllerOff,
	bHomeCompleted 		:= bHomeCompleted,
	Axis 				:= Axis,
	MasterAxis 			:= MasterAxis
 );
END_ACTION

ACTION A_AxisMoveManual:

(* Move axis manual *)
fbMoveManual(
	bEnable 		:= bNoEStop
               		    AND bPowerSupplyOn
               		    AND bSafetyOK,
	bCtrlEnabled 	:= bCtrlEnabled
                		AND bMoveRelease,
	etMachineMode 	:= etMachineMode,
	etMachineState 	:= etMachineState,
	bReset 			:= bConfirmAlarm,
	bMovePlus 		:= bTipPlus,
	bMoveMinus 		:= bTipMinus,
	lrTipDistance 	:= lrTipDistance,
	bLimitMax 		:= bHardLimitMaxExceeded
			      	 	OR bSoftLimitMaxExceeded ,
	bLimitMin 		:= bHardLimitMinExceeded
			      		OR bSoftLimitMinExceeded,
	bPlusRelease 	:= bPlusRelease,
	bMinusRelease 	:= bMinusRelease,
	lrVelocity 		:= SEL(NOT bReferenced, lrManualVelocity, lrVelocityNoRef),
	lrAcceleration 	:= lrAcceleration,
	lrDeceleration 	:= lrDeceleration,
	lrJerk 			:= lrJerk,
	tControllerOff 	:= tControllerOff,
	bHomeCompleted 	:= bHomeCompleted,
	Axis 			:= Axis,
	MasterAxis		:= MasterAxis
);

bSafetyLock := fbMoveManual.bMovePlus
                		OR fbMoveManual.bMoveMinus;
END_ACTION

ACTION A_AxisTerminalDiag:

(*Axis terminal diagnosis *)
fbTerminalDiagnosis(
	stTerminalState := Drive.stTerminalState,
	sTerminalStatus => sTerminalStatus
);

bErrorTerminal := NOT fbTerminalDiagnosis.bTerminalOK;
END_ACTION

END_FUNCTION_BLOCK

// ---- POUs/Machine/Group_0500 - Transport/Gr05Control/Gr05Units/FB_Gr05CylinderClamp.TcPOU
FUNCTION_BLOCK FB_Gr05CylinderClamp
(*

The function block used to lock/unlock welding head.

Constructor: 		Patryk Panylo
Company:			E. Riexinger GmbH
Date:				28.04.2015
Version:			1.00

Date:			Revision:		Who:				Comment
dd.mm.yyyy		x.xx			Initials			comment

*)
VAR_INPUT
	(* Input variables / Eingang Variablen *)
	etMachineMode				:ET_MachineMode;			(* Machine mode *)
	etMachineState				:ET_MachineState;			(* Machine state *)
	bAirPressureOK				:BOOL;						(* Air pressure OK *)
	bSafetyOk					:BOOL;						(* Safety Ok *)
	bOpened						:BOOL;						(* Opened *)
	bClosed						:BOOL;						(* Closed *)
	bOpenRelease				:BOOL;						(* Release open *)
	bCloseRelease				:BOOL;						(* Release close *)
	bHandOpen					:BOOL;						(* Hand open *)
	bHandClose					:BOOL;						(* Hand close *)
	bAutoOpen					:BOOL;						(* Auto open *)
	bAutoClose					:BOOL;						(* Auto close *)
	bExtAutoCtrlEn				:BOOL;						(* Enable external auto control *)
	bExtOpen					:BOOL;						(* External open *)
	bExtClose					:BOOL;						(* External close *)
	bControlOff					:BOOL;						(* TRUE - controle off *)
	bControlStateOn				:BOOL;						(* Control with input state *)
	bValveOff					:BOOL;						(* Valve off *)
	bConfirmAlarm				:BOOL;						(* Confirm alarm *)
	tTimeOut					:TIME := T#6S;				(* TimeOut *)
END_VAR
VAR_OUTPUT
	(* Output variables / Ausgang Variablen *)
	bOpen						:BOOL;						(* Open *)
	bClose						:BOOL;						(* Close *)
	bErrorOpen					:BOOL;						(* Error open *)
	bErrorClose					:BOOL;						(* Error close *)
END_VAR
VAR_IN_OUT
	(* Input Output variables / Ausgang Variablen *)
	bHomeCompleted				:BOOL;						(* Home completed *)
END_VAR
VAR
	(* Enummerations *)

	(* Variables *)

	(* References *)

	(* Interfaces *)

	(* Instances *)
	fbCylinder					:FB_Cylinder;
	fbCylinderOpened				:FB_SignalHandlingDelay;
	fbCylinderClosed				:FB_SignalHandlingDelay;
	fbCylinderOpenRelease		:FB_SignalHandlingDelay;
	fbCylinderCloseRelease		:FB_SignalHandlingDelay;
	fbExtOpen					:FB_SignalHandlingEdge;
	fbExtClose					:FB_SignalHandlingEdge;

END_VAR


(* Control clamp cylinder *)

fbCylinderOpened(
	bEnable := TRUE,
	bIn := bOpened,
	tDelay := t#0ms
);

fbCylinderClosed(
	bEnable := TRUE,
	bIn := bClosed,
	tDelay := 	t#3s
);

fbCylinderOpenRelease(
	bEnable := TRUE,
	bIn := bOpenRelease,
	tDelay :=t#0ms
);

fbCylinderCloseRelease(
	bEnable := TRUE,
	bIn := bCloseRelease,
	tDelay := t#0ms
);

fbExtOpen(
	bEnable := TRUE,
	bIn := bExtOpen,
	tDelay := t#0ms
);

fbExtClose(
	bEnable := TRUE,
	bIn := bExtClose,
	tDelay := t#0ms
);

fbCylinder(
	bEnable := TRUE,
	bAirPressure := bAirPressureOK,
	bSafetyOk := bSafetyOk,
	bReset := bConfirmAlarm,
	bAutoHand := etMachineMode = ET_MachineMode_eHome
			         OR etMachineMode = ET_MachineMode_eStepping
			         OR etMachineMode = ET_MachineMode_eAutomatic,
	bHandBase := bHandOpen OR fbExtOpen.bRisingEdge,
	bHandWork := bHandClose OR fbExtClose.bRisingEdge,
	bAutoBase := SEL(bExtAutoCtrlEn, bAutoOpen, fbExtOpen.bRisingEdge),
	bAutoWork := SEL(bExtAutoCtrlEn, bAutoClose, fbExtClose.bRisingEdge),
	bAtBasePos := fbCylinderOpened.bOut,
	bAtWorkPos := fbCylinderClosed.bOut,
	bBaseRelease := fbCylinderOpenRelease.bOut,
	bWorkRelease := fbCylinderCloseRelease.bOut,
	bControlStateOn := bControlStateOn,
	bControlOff := bControlOff,
	bValveOff := bValveOff,
	bValveErrOff := FALSE,
	bErrorOff := FALSE,
	tTimeOut := tTimeOut + fbCylinderClosed.tDelay,
	bHomeCompleted := bHomeCompleted,
	bMoveToBase => bOpen,
	bMoveToWork => bClose
);

A_Alarm();

ACTION A_Alarm:

bErrorClose := fbCylinder.bError
			AND (fbCylinder.udnErrorNo = 1
				   OR fbCylinder.udnErrorNo = 2
				   OR fbCylinder.udnErrorNo = 5);

bErrorOpen := fbCylinder.bError
			 AND (fbCylinder.udnErrorNo = 3
			       	    OR fbCylinder.udnErrorNo = 4
			       	    OR fbCylinder.udnErrorNo = 5);
END_ACTION

END_FUNCTION_BLOCK

// ---- POUs/Tc2 Objects/Automation/Cylinder/FB_Cylinder.TcPOU
FUNCTION_BLOCK FB_Cylinder
(*
Base class of cylinder.
Cylinder control two directions with handshake.

Constructor: 		Patryk Panylo
Company:		E. Riexinger GmbH
Date:			06.03.2013
Version:			1.00

Date:			Revision:		Who:				Comment
10.30.2013		.02				PPA					Error diagnose off
10.02.2015		.03				PPA					Move in manual in spite of error
13.05.2016		.04				PPA					Valve Off if came limit imput, Control outputs dependent on input state
10.09.2019		.05				PPA					Safety
*)
VAR_INPUT
	(* Input variables / Eingang Variablen *)
	bEnable						:BOOL;			(* Signal FB enable *)
	bAirPressure					:BOOL;			(* Signal air pressure *)
	bSafetyOk					:BOOL;			(* Safety OK  *)
	bReset						:BOOL;			(* Signal reset *)
	bAutoHand					:BOOL;			(* Auto := TRUE, Hand := FALSE *)
	bHandBase					:BOOL;			(* Move hand to base position *)
	bHandWork					:BOOL;			(* Move hand to work position *)
	bAutoBase					:BOOL;			(* Move auto to base position *)
	bAutoWork					:BOOL;			(* Move auto to work position *)
	bAtBasePos					:BOOL;			(* At base position *)
	bAtWorkPos					:BOOL;			(* At work position *)
	bBaseRelease				:BOOL;			(* Base position release *)
	bWorkRelease				:BOOL;			(* Work position release *)
	bControlStateOn				:BOOL;			(* TRUE - control with input state *)
	bControlOff					:BOOL;			(* TRUE - controle off *)
	bValveOff					:BOOL;			(* TRUE -  valve off with limit input *)
	bValveErrOff					:BOOL;			(* TRUE -  valve off if error *)
	bErrorOff						:BOOL;			(* TRUE - error diagnose off *)
	tTimeOut						:TIME := T#5s;	(* TimeOut *)
END_VAR
VAR_OUTPUT
	(* Output variables / Ausgang Variablen *)
	bMoveToBase				:BOOL;			(* Move to base position *)
  	bMoveToWork				:BOOL;			(* Move to work position *)
	bEndBase					:BOOL;			(* Base position reached *)
  	bEndWork					:BOOL;			(* Work position reached *)
 	bNoEndPos					:BOOL;			(* End position not reached *)
	bSafetyLock					:BOOL;			(* Lock safety because of moving *)
	bError						:BOOL;			(* Error *)
	udnErrorNo					:UDINT;			(* Error number *)
	sErrorMsg					:STRING; 		(* Error message *)
END_VAR
VAR_IN_OUT
	(* Input Output variables / Ausgang Variablen *)
	bHomeCompleted				:BOOL;			(* Home completed *)
END_VAR
VAR
	(* Enummerations *)

	(* Variables *)
	bTargetBase					:BOOL;
	bTargetWork					:BOOL;

	bFirstTime					:BOOL;
	(* References *)

	(* Interfaces *)

	(* Instances *)
	rtHandBase					:R_TRIG;
	rtHandWork					:R_TRIG;
	rtAutoBase					:R_TRIG;
	rtAutoWork					:R_TRIG;

 	tonWatchDog					:TON;
END_VAR

IF NOT bEnable
THEN
	bMoveToBase := FALSE;			(* Move to base position *)
  	bMoveToWork := FALSE;			(* Move to work position *)
	bEndBase := FALSE;				(* Base position reached *)
  	bEndWork := FALSE;				(* Work position reached *)
	bError := FALSE;
	udnErrorNo := 0;					(* Error number *)
	sErrorMsg := ''; 					(* Error message *)
	tonWatchDog(IN := FALSE);
	bFirstTime := FALSE;
	RETURN;
END_IF


IF NOT bFirstTime
THEN
	bMoveToBase := FALSE;			(* Move to base position *)
  	bMoveToWork := FALSE;			(* Move to work position *)
	bTargetBase := FALSE;
	bTargetWork := FALSE;
	bEndBase := FALSE;				(* Base position reached *)
  	bEndWork := FALSE;				(* Work position reached *)
	bFirstTime := TRUE;
	RETURN;
END_IF;

(* Air pressure ok / Luftdruck ok *)
IF NOT bAirPressure
THEN
	rtHandBase(CLK:= FALSE);
	rtHandWork(CLK:= FALSE);
	bSafetyLock := FALSE;
	RETURN;
END_IF;

(* Safety lock *)
bSafetyLock := bHandBase
			  OR bHandWork;

A_SetInputs();
A_ChkOpMode();
A_SetOutputs();
A_Status();

ACTION A_ChkOpMode:

(* Check operating mode *)
IF bAutoHand					(* Automatic *)
THEN
	IF rtAutoBase.Q
	     AND NOT bError
	THEN
		bTargetBase := TRUE;
		bTargetWork := FALSE;
	END_IF;

	IF rtAutoWork.Q
 	     AND NOT bError
	THEN
		bTargetBase := FALSE;
		bTargetWork := TRUE;
	END_IF;

ELSE						(* Manual *)
	IF rtHandBase.Q
	    AND bBaseRelease
	    (* AND NOT bError *)
	THEN
		bTargetBase := TRUE;
		bTargetWork := FALSE;
	END_IF;

	IF rtHandWork.Q
	    AND bWorkRelease
	    (* AND NOT bError *)
	THEN
		bTargetBase := FALSE;
		bTargetWork := TRUE;
	END_IF

END_IF;
END_ACTION

ACTION A_SetInputs:

(* Check inputs  *)
rtHandBase(CLK:= bHandBase AND bSafetyOk);
rtHandWork(CLK:= bHandWork AND bSafetyOk);
rtAutoBase(CLK:= bAutoBase AND bBaseRelease AND bSafetyOk);
rtAutoWork(CLK:= bAutoWork AND bWorkRelease AND bSafetyOk);
END_ACTION

ACTION A_SetOutputs:

(* Set outputs move to base position  *)
IF bBaseRelease
     OR bAtBasePos
THEN
	IF  bTargetBase
	     AND NOT bMoveToBase
	THEN
		bMoveToBase := TRUE;
		bMoveToWork := FALSE;
		tonWatchDog(IN := FALSE);
	END_IF;

ELSE
	IF bTargetBase
	     AND  bMoveToBase
	THEN
		bMoveToBase := FALSE;

		IF NOT bAutoHand
		THEN
			bTargetBase := FALSE;
		END_IF;

	END_IF;
END_IF;

(* Set outputs move to work position  *)
IF bWorkRelease
    OR bAtWorkPos
THEN
	IF  bTargetWork
	     AND NOT bMoveToWork
	THEN
		bMoveToBase := FALSE;
		bMoveToWork := TRUE;
		tonWatchDog(IN := FALSE);
	END_IF;

ELSE
	IF bTargetWork
	     AND  bMoveToWork
	THEN
		bMoveToWork := FALSE;

		IF NOT bAutoHand
		THEN
			bTargetWork := FALSE;
		END_IF;

	END_IF;
END_IF;

IF NOT bAutoHand
    AND (bMoveToBase
         	       OR bMoveToWork)
THEN
	bHomeCompleted := FALSE;
END_IF;
END_ACTION

ACTION A_Status:

(* Error reset *)
IF bReset
     AND bError
THEN
	udnErrorNo := 0;					(* Error number *)
	sErrorMsg := ''; 					(* Error message *)
	tonWatchDog(IN := FALSE);
END_IF;

(* Timer starts when cylinder is not  in base and work position *)
tonWatchDog(IN := NOT bErrorOff
				 AND (
					(bMoveToWork AND NOT bAtWorkPos)
				   	OR (bMoveToBase AND NOT bAtBasePos)
				   	OR (NOT bAtBasePos AND NOT bAtWorkPos)
				   	OR (bAtBasePos AND bAtWorkPos)),
			PT := tTimeOut);

(* Error if cylinder does not reach base or work position*)
IF tonWatchDog.Q 
   AND NOT bError
THEN
	IF bMoveToWork
	THEN
		IF NOT bAtWorkPos AND NOT bAtBasePos
		THEN
			udnErrorNo := 1; 								(* Set error number *)
			sErrorMsg := 'Work position not reached';
		ELSIF NOT bAtWorkPos AND bAtBasePos
		THEN
			udnErrorNo := 2; 								(* Set error number *)
			sErrorMsg := 'Not move in work position';
		ELSIF bAtWorkPos AND bAtBasePos
		THEN
			udnErrorNo := 5; 									(* Set error number *)
			sErrorMsg := 'Both position reached';
		END_IF
	ELSIF bMoveToBase
	THEN
		IF NOT bAtWorkPos AND NOT bAtBasePos
		THEN
			udnErrorNo := 3; 								(* Set error number *)
			sErrorMsg := 'Base position not reached';
		ELSIF bAtWorkPos AND NOT bAtBasePos
		THEN
			udnErrorNo := 4; 								(* Set error number *)
			sErrorMsg := 'Not move in base position';
		ELSIF bAtWorkPos AND bAtBasePos
		THEN
			udnErrorNo := 5; 									(* Set error number *)
			sErrorMsg := 'Both position reached';
		END_IF
	ELSIF bAtWorkPos AND bAtBasePos
	THEN
		udnErrorNo := 5; 									(* Set error number *)
		sErrorMsg := 'Both position reached';
	END_IF
END_IF

bError := udnErrorNo <> 0;


(* End base position reached  *)
bEndBase := bAtBasePos
		        AND NOT bAtWorkPos
		        AND NOT bError;

(* End wrok position reached  *)
bEndWork := NOT bAtBasePos
		        AND bAtWorkPos
		        AND NOT bError;

(* End position not reached *)
IF bTargetBase
THEN
	bNoEndPos := NOT bAtBasePos;

ELSIF bTargetWork
THEN
	bNoEndPos :=  NOT bAtWorkPos;

ELSE
	bNoEndPos := FALSE;
END_IF


(* Valve off if error  *)
IF bError
     AND (bMoveToBase OR bMoveToWork)
     AND bValveErrOff
THEN
	bMoveToBase := FALSE;
	bMoveToWork := FALSE;
	bTargetBase := FALSE;
	bTargetWork := FALSE;
END_IF;

(* Control with input state *)
IF bControlStateOn
THEN
	IF bAutoHand					(* Automatic *)
	THEN
		IF NOT bAutoBase
		THEN
			bMoveToBase := FALSE;
			bTargetBase := FALSE;
		END_IF

		IF NOT bAutoWork
		THEN
			bMoveToWork := FALSE;
			bTargetWork := FALSE;
		END_IF
	
	ELSE						(* Manual *)
		IF NOT bHandBase
		THEN
			bMoveToBase := FALSE;
			bTargetBase := FALSE;
		END_IF

		IF NOT bHandWork
		THEN
			bMoveToWork := FALSE;
			bTargetWork := FALSE;
		END_IF
	
	END_IF;
END_IF

(* Check control off *)
IF bControlOff
    AND (
		bMoveToBase OR bMoveToWork
		OR bTargetBase OR bTargetWork
	      )
THEN
	bMoveToBase := FALSE;
	bMoveToWork := FALSE;
	bTargetBase := FALSE;
	bTargetWork := FALSE;
END_IF

(* Check valve off *)
IF bValveOff
THEN
	IF bAtBasePos
	    AND (bMoveToBase OR bTargetBase)
	THEN
		bMoveToBase := FALSE;
		bTargetBase := FALSE;

	ELSIF bAtWorkPos
	    	   AND (bMoveToWork OR bTargetWork)
	THEN
		bMoveToWork := FALSE;
		bTargetWork := FALSE;
	END_IF
END_IF
END_ACTION

END_FUNCTION_BLOCK

// ---- POUs/Machine/Group_0500 - Transport/Gr05Control/Gr05Units/FB_Gr05CylinderPos.TcPOU
FUNCTION_BLOCK FB_Gr05CylinderPos
(*

The function block used to control position cylinder.

Constructor: 		Patryk Panylo
Company:		E. Riexinger GmbH
Date:			28.04.2015
Version:			1.00

Date:			Revision:		Who:				Comment
dd.mm.yyyy		x.xx			Initials			comment

*)
VAR_INPUT
	(* Input variables / Eingang Variablen *)
	bEnable						:BOOL;															(* Function block enable *)
	etMachineMode				:ET_MachineMode;												(* Machine mode *)
	etMachineState				:ET_MachineState;												(* Machine state *)
	bNoEStop					:BOOL;															(* No ermergency Stop / Keine Notaus *)
	bSafetyOK					:BOOL;															(* Safety ok / Sicherheit i.o *)
	bAirPressureOK				:BOOL;															(* Air pressure OK *)
	bExeMoveAbs				:BOOL;															(* Execute move absolut *)
	lrTargetPosition				:LREAL;															(* Absolute target position *)
	arbInBase					:ARRAY[1..ungGr05CylinderPosMaxNo] OF BOOL;						(* In base position *)
	arbInWork					:ARRAY[1..ungGr05CylinderPosMaxNo] OF BOOL;						(* In work position *)
	arbMoveToBaseRelease		:ARRAY[1..ungGr05CylinderPosMaxNo] OF BOOL;						(* Release move to base *)
	arbMoveToWorkRelease		:ARRAY[1..ungGr05CylinderPosMaxNo] OF BOOL;						(* Release move to work *)
	arbHandMoveToBase			:ARRAY[1..ungGr05CylinderPosMaxNo] OF BOOL;						(* Hand move to base *)
	arbHandMoveToWork			:ARRAY[1..ungGr05CylinderPosMaxNo] OF BOOL;						(* Hand move to work *)
	lrPosOffset					:LREAL;															(* Position offset *)
	lrOriginShiftPos				:LREAL;															(* Origin shift position *)
	etDirection					:ET_MC_Direction;													(* Direction: -1 Negative, +1 Positive *)
	usnCodingType				:USINT;
	bControlStateOn				:BOOL;															(* Control with input state *)
	bControlOff					:BOOL;															(* Controle off *)
	bValveOff					:BOOL;															(* Valve off *)
	bConfirmAlarm				:BOOL;															(* Confirm alarm *)
	tTimeOut						:TIME := t#6s;														(* TimeOut *)
END_VAR
VAR_OUTPUT
	(* Output variables / Ausgang Variablen *)
	bCtrlEnabled					:BOOL;						(* Controller enabled *)
	lrActPosition					:LREAL;															(* Actual position [mm] *)
	arbMoveToBase				:ARRAY[1..ungGr05CylinderPosMaxNo] OF BOOL;						(* Move to base *)
	arbMoveToWork				:ARRAY[1..ungGr05CylinderPosMaxNo] OF BOOL;						(* Move to work *)
	arbErrorMoveToBase			:ARRAY[1..ungGr05CylinderPosMaxNo] OF BOOL;						(* Error move to base *)
	arbErrorMoveToWork			:ARRAY[1..ungGr05CylinderPosMaxNo] OF BOOL;						(* Error move to work *)
END_VAR
VAR_IN_OUT
	(* Input Output variables / Ausgang Variablen *)
	bHomeCompleted				:BOOL;						(* Home completed *)
END_VAR
VAR
	(* Enummerations *)

	(* Variables *)
	unCylinderPosIdx				:UINT;						(* Position cylinder index *)

	(* References *)

	(* Interfaces *)

	(* Instances *)
	fbCylinderPos				:ARRAY[1..ungGr05CylinderPosMaxNo] OF FB_CylinderPos;
	fbMoveAbs					:FB_CylinderPos_MoveAbsolut;
END_VAR


(* Control position cylinder cylinder *)
(*
lrRefPos := TAN(ABS(lrAngle)) * (lrRadius + lrSafetyDistance);
*)

fbMoveAbs(
	bEnable := bEnable,
	bNoEStop := bNoEStop,
	bLightCurtainOK := bSafetyOK,
	bAirPressure := bAirPressureOK,
	bExecute := bExeMoveAbs,
	lrPosition := lrTargetPosition,
	lrPosOffset := lrPosOffset,
	lrOriginShiftPos := lrOriginShiftPos,
	etDirection := etDirection,
	usnCodingType := usnCodingType,
	lrActPosition => lrActPosition
);

FOR unCylinderPosIdx := 1 TO ungGr05CylinderPosMaxNo
DO

	fbCylinderPos[unCylinderPosIdx](
		etMachineMode := etMachineMode,
		etMachineState := etMachineState,
		bAirPressureOK := bAirPressureOK,
		bSafetyOK := bSafetyOK,
		bInBase := arbInBase[unCylinderPosIdx],
		bInWork := arbInWork[unCylinderPosIdx],
		bMoveToBaseRelease := TRUE,
		bMoveToWorkRelease := TRUE,
		bHandMoveToBase := arbHandMoveToBase[unCylinderPosIdx],
		bHandMoveToWork := arbHandMoveToWork[unCylinderPosIdx],
		bAutoMoveToBase := fbMoveAbs.arbToBase[unCylinderPosIdx],
		bAutoMoveToWork := fbMoveAbs.arbToWork[unCylinderPosIdx],
		bConfirmAlarm := bConfirmAlarm,
		bControlStateOn := bControlStateOn,
		bControlOff := bControlOff,
		bValveOff := bValveOff,
		bValveErrOff := FALSE,
		bErrorOff := FALSE,
		tTimeOut := t#6s,
		bHomeCompleted := bHomeCompleted,
		bMoveToBase => arbMoveToBase[unCylinderPosIdx],
		bMoveToWork => arbMoveToWork[unCylinderPosIdx]
	);

	fbMoveAbs.arbInBase[unCylinderPosIdx] := fbCylinderPos[unCylinderPosIdx].fbCylinderPos.bEndBase;
	fbMoveAbs.arbInWork[unCylinderPosIdx] := fbCylinderPos[unCylinderPosIdx].fbCylinderPos.bEndWork;
	fbMoveAbs.arbInError [unCylinderPosIdx] := fbCylinderPos[unCylinderPosIdx].fbCylinderPos.bError;

END_FOR

bCtrlEnabled := bNoEStop
			   AND bSafetyOK
			   AND bAirPressureOK;

A_Alarm();

ACTION A_Alarm:

FOR unCylinderPosIdx := 1 TO ungGr05CylinderPosMaxNo
DO

	arbErrorMoveToBase[unCylinderPosIdx] := fbCylinderPos[unCylinderPosIdx].bErrorMoveToBase;
	arbErrorMoveToWork[unCylinderPosIdx] := fbCylinderPos[unCylinderPosIdx].bErrorMoveToWork;

END_FOR
END_ACTION

END_FUNCTION_BLOCK

// ---- POUs/Machine/Group_0500 - Transport/Gr05Control/Gr05Units/FB_Gr05Slide.TcPOU
FUNCTION_BLOCK FB_Gr05Slide
(*

The function block used to control slide.

Constructor: 		Patryk Panylo
Company:		E. Riexinger GmbH
Date:			28.04.2015
Version:			1.00

Date:			Revision:		Who:				Comment
dd.mm.yyyy		x.xx			Initials			comment

*)
VAR_INPUT
	(* Input variables / Eingang Variablen *)
	bEnable						:BOOL;						(* FB enable *)
	etMachineMode				:ET_MachineMode;			(* Machine mode *)
	etMachineState				:ET_MachineState;			(* Machine state *)
	bAirPressureOK				:BOOL;						(* Air pressure OK *)
	bSafetyOk					:BOOL;						(* Safety Ok *)
	bInBase						:BOOL;						(* In base position *)
	bInWork						:BOOL;						(* In work position *)
	bMoveToBaseRelease		:BOOL;						(* Release move to base *)
	bMoveToWorkRelease		:BOOL;						(* Release move to work *)
	bHandMoveToBase			:BOOL;						(* Hand move to base *)
	bHandMoveToWork			:BOOL;						(* Hand move to work *)
	bAutoMoveToBase			:BOOL;						(* Auto move to base *)
	bAutoMoveToWork			:BOOL;						(* Auto move to work *)
	bControlStateOn				:BOOL;						(* Control with input state *)
	bControlOff					:BOOL;						(* Controle off *)
	bValveOff					:BOOL;						(* Valve off *)
	bConfirmAlarm				:BOOL;						(* Confirm alarm *)
	tTimeOut						:TIME := t#6s;					(* TimeOut *)
END_VAR
VAR_OUTPUT
	(* Output variables / Ausgang Variablen *)
	bMoveToBase				:BOOL;						(* Move to base *)
	bMoveToWork				:BOOL;						(* Move to work *)
	bErrorMoveToBase			:BOOL;						(* Error move to base *)
	bErrorMoveToWork			:BOOL;						(* Error move to work *)
END_VAR
VAR_IN_OUT
	(* Input Output variables / Ausgang Variablen *)
	bHomeCompleted				:BOOL;						(* Home completed *)
END_VAR
VAR
	(* Enummerations *)

	(* Variables *)

	(* References *)

	(* Interfaces *)

	(* Instances *)
	fbCylinder					:FB_Cylinder;
	fbCylinderAtBasePos			:FB_SignalHandlingDelay;
	fbCylinderAtWorkPos			:FB_SignalHandlingDelay;
	fbCylinderBaseRelease		:FB_SignalHandlingDelay;
	fbCylinderWorkRelease		:FB_SignalHandlingDelay;

END_VAR


IF NOT bEnable								(* Signal FB enable *)
THEN

	RETURN;
END_IF

(* Control slide cylinder *)

fbCylinderAtBasePos(
	bEnable := TRUE,
	bIn := bInBase,
	tDelay := t#0ms
);

fbCylinderAtWorkPos(
	bEnable := TRUE,
	bIn := bInWork,
	tDelay := t#0ms
);

fbCylinderBaseRelease(
	bEnable := TRUE,
	bIn := bMoveToBaseRelease,
	tDelay :=t#0ms
);

fbCylinderWorkRelease(
	bEnable := TRUE,
	bIn := bMoveToWorkRelease,
	tDelay := t#0ms
);

fbCylinder(
	bEnable := TRUE,
	bAirPressure := bAirPressureOK,
	bSafetyOk := bSafetyOk,
	bReset := bConfirmAlarm,
	bAutoHand := etMachineMode = ET_MachineMode_eHome
			         OR etMachineMode = ET_MachineMode_eStepping
			         OR etMachineMode = ET_MachineMode_eAutomatic,
	bHandBase := bHandMoveToBase,
	bHandWork := bHandMoveToWork,
	bAutoBase := bAutoMoveToBase,
	bAutoWork := bAutoMoveToWork,
	bAtBasePos := fbCylinderAtBasePos.bOut,
	bAtWorkPos := fbCylinderAtWorkPos.bOut,
	bBaseRelease := fbCylinderBaseRelease.bOut,
	bWorkRelease := fbCylinderWorkRelease.bOut,
	bControlStateOn := bControlStateOn,
	bControlOff := bControlOff,
	bValveOff := bValveOff,
	bValveErrOff := FALSE,
	bErrorOff := FALSE,
	tTimeOut := tTimeOut,
	bHomeCompleted := bHomeCompleted,
	bMoveToBase => bMoveToBase,
	bMoveToWork => bMoveToWork
);

A_Alarm();

ACTION A_Alarm:

bErrorMoveToWork := fbCylinder.bError
					AND (fbCylinder.udnErrorNo = 1
					     OR fbCylinder.udnErrorNo = 2
					     OR fbCylinder.udnErrorNo = 5);

bErrorMoveToBase := fbCylinder.bError
					 AND (fbCylinder.udnErrorNo = 3
					       OR fbCylinder.udnErrorNo = 4
					       OR fbCylinder.udnErrorNo = 5);
END_ACTION

END_FUNCTION_BLOCK

// ---- POUs/Machine/Group_0500 - Transport/Gr05Control/Gr05Units/FB_Gr05RemovalBand.TcPOU
FUNCTION_BLOCK FB_Gr05RemovalBand
(*

The function block used to remove parts.

Constructor: 		Patryk Panylo
Company:		E. Riexinger GmbH
Date:			28.04.2015
Version:			1.00

Date:			Revision:		Who:				Comment
dd.mm.yyyy		x.xx			Initials			comment

*)
VAR_INPUT
	(* Input variables / Eingang Variablen *)
	etMachineMode				:ET_MachineMode;			(* Machine mode *)
	etMachineState				:ET_MachineState;			(* Machine state *)
	bNoEStop					:BOOL;						(* No ermergency Stop / Keine Notaus *)
	bPowerSupplyOn				:BOOL;						(* Power supply on / Leitung eingeschaltet *)
	bSafetyOK					:BOOL;						(* Safety ok / Sicherheit i.o *)
	bInPlusLimit					:BOOL;						(* In plus limit *)
	bInMinusLimit					:BOOL;						(* In minus limit *)
	bMoveToPlusRelease			:BOOL;						(* Release move to plus *)
	bMoveToMinusRelease		:BOOL;						(* Release move to minus *)
	bHandMoveToPlus			:BOOL;						(* Hand move to pluse *)
	bHandMoveToMinus			:BOOL;						(* Hand move to minus *)
	bAutoMoveToPlus			:BOOL;						(* Auto move to plus *)
	arbAutoMoveToMinus			:ARRAY[1..2] OF BOOL;		(* Auto move to minus *)
	bConfirmAlarm				:BOOL;						(* Confirm alarm *)
	tTimeOut						:TIME := t#6s;					(* TimeOut *)
END_VAR
VAR_OUTPUT
	(* Output variables / Ausgang Variablen *)
	bMoveToPlus				:BOOL;						(* Move to plus *)
	bMoveToMinus				:BOOL;						(* Move to minus *)
	bErrorMoveToPlus			:BOOL;						(* Error move to plus *)
	bErrorMoveToMinus			:BOOL;						(* Error move to minus *)
END_VAR
VAR_IN_OUT
	(* Input Output variables / Ausgang Variablen *)
	bHomeCompleted				:BOOL;						(* Home completed *)
END_VAR
VAR
	(* Enummerations *)

	(* Variables *)

	(* References *)

	(* Interfaces *)

	(* Instances *)
	fbMotor					:FB_Motor;
	fbMotorAtPlusLimit			:FB_SignalHandlingDelay;
	fbMotorAtMinusLimit		:FB_SignalHandlingDelay;
	fbMotorPlusRelease		:FB_SignalHandlingDelay;
	fbMotorMinusRelease		:FB_SignalHandlingDelay;
	tofAutoMoveToMinus		:TOF;
END_VAR


(* Control removal band motor *)

fbMotorAtPlusLimit(
	bEnable := TRUE,
	bIn := bInPlusLimit,
	tDelay := t#0ms
);

fbMotorAtMinusLimit(
	bEnable := TRUE,
	bIn := bInMinusLimit,
	tDelay := t#0ms
);

fbMotorPlusRelease(
	bEnable := TRUE,
	bIn := bMoveToPlusRelease,
	tDelay :=t#0ms
);

fbMotorMinusRelease(
	bEnable := TRUE,
	bIn := bMoveToMinusRelease,
	tDelay := t#0ms
);

tofAutoMoveToMinus(
	IN := arbAutoMoveToMinus[1]
		OR arbAutoMoveToMinus[2],				(* Auto move to minus *)
	PT := t#0s,
);

fbMotor(
	bEnable := TRUE,
	bNoEmergencyStop := bNoEStop
						AND bSafetyOK,
	bVoltageOK := bPowerSupplyOn,
	bReset := bConfirmAlarm,
	bAutoHand := etMachineMode = ET_MachineMode_eHome
			         OR etMachineMode = ET_MachineMode_eStepping
			         OR etMachineMode = ET_MachineMode_eAutomatic,
	bHandPlus := bHandMoveToPlus,
	bHandMinus := bHandMoveToMinus,
	bAutoPlus := bAutoMoveToPlus,
	bAutoMinus := tofAutoMoveToMinus.Q,
	bAtPlusLimit := fbMotorAtPlusLimit.bOut,
	bAtMinusLimit := fbMotorAtMinusLimit.bOut,
	bPlusRelease := fbMotorPlusRelease.bOut,
	bMinusRelease := fbMotorMinusRelease.bOut,
	bSyncPlus := FALSE,
	bSyncMinus := FALSE,
	bSyncOn := FALSE,
	bControlOff := NOT bHandMoveToMinus
				AND NOT tofAutoMoveToMinus.Q,
	tControlOff := t#1s500ms,
	bMotorCtrlErrOff := FALSE,
	bErrorOff := TRUE,
	tSyncTimeOut := ,
	tConTimeOut := ,
	tCtrlTimeOut := tTimeOut,
	bHomeCompleted := bHomeCompleted,
	bMoveToPlus => bMoveToPlus,
	bMoveToMinus => bMoveToMinus
);

A_Alarm();

ACTION A_Alarm:

bErrorMoveToPlus := fbMotor.bError
					AND (fbMotor.udnErrorNo = 1
					     OR fbMotor.udnErrorNo = 2
					     OR fbMotor.udnErrorNo = 5);

bErrorMoveToMinus := fbMotor.bError
					 AND (fbMotor.udnErrorNo = 3
					       OR fbMotor.udnErrorNo = 4
					       OR fbMotor.udnErrorNo = 5);
END_ACTION

END_FUNCTION_BLOCK

// ---- POUs/Tc2 Objects/Automation/MotorOnOff/FB_Motor.TcPOU
FUNCTION_BLOCK FB_Motor
(*
Base class of motor.
Motor controls with handshake.

Constructor: 		Patryk Panylo
Company:		E. Riexinger GmbH
Date:			19.04.2013
Version:			1.00

Date:			Revision:		Who:				Comment
22.04.2013		.01				PPA					Motor binary synchronization
03.05.2013		.02				PPA					Condition monitoring
30.10.2013		.03				PPA					Error diagnose off
05.12.2016		.04				PPA					External alarm
*)
VAR_INPUT
	bEnable					:BOOL;
	bNoEmergencyStop		:BOOL;			(* Emergency stop / NotAus *)
	bVoltageOK				:BOOL;			(* Voltage OK *)
	bExtAlarm				:BOOL;			(* External alarm *)
	bReset					:BOOL;
	bAutoHand				:BOOL;			(* Auto := TRUE, Hand := FALSE *)
	bHandPlus				:BOOL;
	bHandMinus				:BOOL;
	bAutoPlus				:BOOL;
	bAutoMinus				:BOOL;
	bAtPlusLimit				:BOOL;			(* At position limit plus *)
	bAtMinusLimit				:BOOL;			(* At position limit minus *)
	bPlusRelease			:BOOL;			(* Plus position release *)
	bMinusRelease			:BOOL;			(* Minus position release *)
	bSyncPlus				:BOOL;			(* Synchronization in plus direction *)
	bSyncMinus				:BOOL;			(* Synchronization in minus direction *)
	bSyncOn					:BOOL;			(* TRUE - synchronization*)
	bControlOff				:BOOL;			(* TRUE - controle off *)
	tControlOff				:TIME;			(* Time > 0 delay to control off *)
	bMotorCtrlErrOff			:BOOL;			(* TRUE -  motor off if error *)
	bErrorOff					:BOOL;			(* TRUE - error diagnose off *)
	tSyncTimeOut			:TIME := T#2s;	(* Synchronization TimeOut *)
	tConTimeOut				:TIME := T#500ms;	(* Condition TimeOut *)
	tCtrlTimeOut				:TIME := T#10s;	(* Control TimeOut *)
END_VAR
VAR_OUTPUT
	bMoveToPlus			:BOOL;			(* Move to plus direction *)
  	bMoveToMinus			:BOOL;			(* Move to minus direction *)
	bLimitPlus				:BOOL;			(* Limit switch plus reached *)
  	bLimitMinus				:BOOL;			(* Limit switch minus reached *)
	bError					:BOOL;
	udnErrorNo				:UDINT;			(* Error number *)
	sErrorMsg				:STRING; 		(* Error message *)
END_VAR
VAR_IN_OUT
	(* Input Output variables / Ausgang Variablen *)
	bHomeCompleted				:BOOL;			(* Home completed *)
END_VAR
VAR
  	tonCtrlWatchDog			:TON;
  	tonConWatchDog			:TON;
  	tonSyncWatchDog		:TON;
	tonControlOff				:TON;
	tonHandPlus				:TON;			(* Delay signal hand plus *)
	tonHandMinus			:TON;			(* Delay signal hand minus *)

	rtHandPlus				:R_TRIG;
	rtHandMinus				:R_TRIG;
	rtAutoPlus				:R_TRIG;
	rtAutoMinus				:R_TRIG;

	rtAutoHand				:R_TRIG;
	ftAutoHand				:F_TRIG;

	bTargetPlus				:BOOL;
	bTargetMinus				:BOOL;

	bFirstTime				:BOOL;

END_VAR
VAR CONSTANT
	tPressDelay 				:TIME := t#200ms;			(* Delay hand signals *)
END_VAR

IF NOT bEnable
THEN
	bMoveToPlus := FALSE;			(* Move to plus direction *)
  	bMoveToMinus := FALSE;			(* Move to minus direction *)
	bLimitPlus := FALSE;				(* Limit switch plus reached *)
  	bLimitMinus := FALSE;				(* Limit switch minus reached *)
	bTargetPlus := FALSE;
	bTargetMinus := FALSE;
	bError := FALSE;
	udnErrorNo := 0;					(* Error number *)
	sErrorMsg := ''; 					(* Error message *)
	tonCtrlWatchDog(IN := FALSE);
	tonConWatchDog(IN := FALSE);
	tonSyncWatchDog(IN := FALSE);
	tonControlOff(IN := FALSE);
	bFirstTime := FALSE;
	RETURN;
END_IF

IF NOT bFirstTime
THEN
	bMoveToPlus := FALSE;			(* Move to plus direction *)
  	bMoveToMinus := FALSE;			(* Move to minus direction *)
	bLimitPlus := FALSE;				(* Limit switch plus reached *)
  	bLimitMinus := FALSE;				(* Limit switch minus reached *)
	bTargetPlus := FALSE;
	bTargetMinus := FALSE;
	bFirstTime := TRUE;
	RETURN;
END_IF

IF NOT bNoEmergencyStop
THEN
	bMoveToPlus := FALSE;			(* Move to plus direction *)
  	bMoveToMinus := FALSE;			(* Move to minus direction *)
	bLimitPlus := FALSE;				(* Limit switch plus reached *)
  	bLimitMinus := FALSE;				(* Limit switch minus reached *)
	bTargetPlus := FALSE;
	bTargetMinus := FALSE;
	tonCtrlWatchDog(IN := FALSE);
	tonSyncWatchDog(IN := FALSE);
	tonControlOff(IN := FALSE);
	RETURN;
END_IF

(* Check inputs  *)
tonHandPlus(IN := bHandPlus AND NOT bHandMinus, PT := tPressDelay);
tonHandMinus(IN := bHandMinus AND NOT bHandPlus, PT := tPressDelay);

rtHandPlus(CLK := tonHandPlus.Q);
rtHandMinus(CLK:= tonHandMinus.Q);

rtAutoPlus(CLK:= bAutoPlus AND bPlusRelease);
rtAutoMinus(CLK:= bAutoMinus AND bMinusRelease);


rtAutoHand(CLK := bAutoHand);
ftAutoHand(CLK := bAutoHand);

IF rtAutoHand.Q
    OR ftAutoHand.Q
THEN
	bMoveToPlus := FALSE;			(* Move to plus direction *)
  	bMoveToMinus := FALSE;			(* Move to minus direction *)
	bTargetPlus := FALSE;
	bTargetMinus := FALSE;
END_IF


(* Check operating mode *)
IF bAutoHand					(* Automatic *)
THEN
	IF rtAutoPlus.Q
	     AND NOT bAtPlusLimit					(* No at position limit plus *)
	     AND NOT bError
	THEN
		bTargetPlus := TRUE;
		bTargetMinus := FALSE;

		tonControlOff(IN := FALSE);

	ELSIF bMoveToPlus
		    AND bAtPlusLimit					(* At position limit plus *)
		    AND NOT bAtMinusLimit				(* No at position limit minus *)
	THEN
		bTargetPlus := FALSE;
		bMoveToPlus := FALSE;				(* Move to plus direction *)

	END_IF

	IF rtAutoMinus.Q
	     AND NOT bAtMinusLimit					(* No at position limit minus *)
 	     AND NOT bError
	THEN
		bTargetPlus := FALSE;
		bTargetMinus := TRUE;

		tonControlOff(IN := FALSE);

	ELSIF bMoveToMinus
		    AND NOT bAtPlusLimit				(* No at position limit plus *)
		    AND bAtMinusLimit					(* At position limit minus *)
	THEN
		bTargetMinus := FALSE;
		bMoveToMinus := FALSE;				(* Move to minus direction *)

	END_IF

ELSE						(* Manual *)

	IF NOT bTargetPlus
	THEN
		IF rtHandPlus.Q
		    AND bPlusRelease
		THEN
			bTargetPlus := TRUE;
			bTargetMinus := FALSE;

			IF bError
			THEN
				bReset  := TRUE;					(*  Error reset *)
			END_IF

		END_IF

	ELSE
		IF NOT bHandPlus
		     OR bAtPlusLimit
		THEN
			bTargetPlus := FALSE;
			bMoveToPlus := FALSE;			(* Move to plus direction *)
		END_IF

	END_IF

	IF NOT bTargetMinus
	THEN
		IF rtHandMinus.Q
		    AND bMinusRelease
		THEN
			bTargetPlus := FALSE;
			bTargetMinus := TRUE;

			IF bError
			THEN
				bReset  := TRUE;					(*  Error reset *)
			END_IF

		END_IF

	ELSE
		IF NOT bHandMinus
		     OR bAtMinusLimit
		THEN
			bTargetMinus := FALSE;
			bMoveToMinus := FALSE;			(* Move to minus direction *)
		END_IF

	END_IF

END_IF

IF NOT bAutoHand
    AND (bMoveToPlus
         	       OR bMoveToMinus)
THEN
	bHomeCompleted := FALSE;
END_IF;

(* Set outputs move to Plus position  *)
IF bPlusRelease								(* Start movement *)
THEN
	IF  bTargetPlus
	     AND NOT bMoveToPlus
	THEN
		bMoveToPlus := TRUE;				(* Move to plus direction *)
		bMoveToMinus := FALSE;
		tonCtrlWatchDog(IN := FALSE);
		tonConWatchDog(IN := FALSE);
		tonSyncWatchDog(IN := FALSE);
	END_IF

ELSE
	IF bTargetPlus							(* Stop movement *)
	     AND  bMoveToPlus
	THEN
		bMoveToPlus := FALSE;

		IF NOT bAutoHand					(* In manual only continue movement *)
		THEN
			bTargetPlus := FALSE;
		END_IF

	END_IF
END_IF

(* Set outputs move to Minus position  *)
IF bMinusRelease								(* Start movment *)
THEN
	IF  bTargetMinus
	     AND NOT bMoveToMinus
	THEN
		bMoveToPlus := FALSE;
		bMoveToMinus := TRUE;				(* Move to minus direction *)
		tonCtrlWatchDog(IN := FALSE);
		tonConWatchDog(IN := FALSE);
		tonSyncWatchDog(IN := FALSE);
	END_IF

ELSE
	IF bTargetMinus							(* Stop movment *)
	     AND  bMoveToMinus
	THEN
		bMoveToMinus := FALSE;

		IF NOT bAutoHand					(* In manual only continue movement *)
		THEN
			bTargetMinus := FALSE;
		END_IF

	END_IF
END_IF


(* Error reset *)
IF bReset
     AND bError
THEN
	udnErrorNo := 0;					(* Error number *)
	sErrorMsg := ''; 					(* Error message *)
	tonCtrlWatchDog(IN := FALSE);
	tonConWatchDog(IN := FALSE);
	tonSyncWatchDog(IN := FALSE);
END_IF;

(* Timer starts when motor is reached plus and minus *)
tonCtrlWatchDog(IN := NOT bErrorOff
				       AND(
					(bMoveToMinus AND NOT bAtMinusLimit)
					OR (bMoveToPlus AND NOT bAtPlusLimit)
				   	OR (NOT bAtPlusLimit AND NOT bAtMinusLimit)
				   	OR (bAtPlusLimit AND bAtMinusLimit)),
			       PT := tCtrlTimeOut);

(* Error if motor does not reach plus or minus limit *)
IF tonCtrlWatchDog.Q
    AND bAutoHand					(* In automatic *)
    AND NOT bError
THEN
	IF bMoveToMinus
	THEN
		IF NOT bAtMinusLimit AND NOT bAtPlusLimit
		THEN
			udnErrorNo := 1; 								(* Set error number *)
			sErrorMsg := 'Minus limit not reached';
		ELSIF NOT bAtMinusLimit AND bAtPlusLimit
		THEN
			udnErrorNo := 2; 								(* Set error number *)
			sErrorMsg := 'Not move in minus limit';
		ELSIF bAtMinusLimit AND bAtPlusLimit
		THEN
			udnErrorNo := 5; 									(* Set error number *)
			sErrorMsg := 'Both position reached';
		END_IF
	ELSIF bMoveToPlus
	THEN
		IF NOT bAtMinusLimit AND NOT bAtPlusLimit
		THEN
			udnErrorNo := 3; 								(* Set error number *)
			sErrorMsg := 'Plus limit not reached';
		ELSIF bAtMinusLimit AND NOT bAtPlusLimit
		THEN
			udnErrorNo := 4; 								(* Set error number *)
			sErrorMsg := 'Not move in plus limit';
		ELSIF bAtMinusLimit AND bAtPlusLimit
		THEN
			udnErrorNo := 5; 									(* Set error number *)
			sErrorMsg := 'Both position reached';
		END_IF
	ELSIF bAtMinusLimit AND bAtPlusLimit
	THEN
		udnErrorNo := 5; 									(* Set error number *)
		sErrorMsg := 'Both position reached';
	END_IF
END_IF

(* Voltage is nok / Spannung nOk *)
IF NOT bVoltageOK
THEN
	IF bMoveToPlus
	     OR bMoveToMinus
	THEN
		bMoveToPlus := FALSE;			(* Move to plus direction *)
	  	bMoveToMinus := FALSE;			(* Move to minus direction *)
		bTargetPlus := FALSE;
		bTargetMinus := FALSE;

		udnErrorNo := 8; 									(* Set error number *)
		sErrorMsg := 'No voltage at motor.';
	END_IF

END_IF

(* Synchronization is nok / Synchronization nOk *)
tonSyncWatchDog(IN := (bMoveToMinus AND NOT bSyncMinus)
					  OR (NOT bMoveToMinus AND bSyncMinus)
				   	  OR (bMoveToPlus AND NOT bSyncPlus)
				  	  OR (NOT bMoveToPlus AND bSyncPlus),
				 PT := tSyncTimeOut);

(* Error if motor not sync plus or minus *)
IF bSyncOn
    AND tonSyncWatchDog.Q
    AND NOT bError
THEN
	IF bMoveToMinus
	THEN
		IF NOT bSyncMinus
		THEN
			udnErrorNo := 10; 									(* Set error number *)
			sErrorMsg := 'Synchronization minus reached';
		END_IF
	ELSIF bMoveToPlus
	THEN
		IF NOT bSyncPlus
		THEN
			udnErrorNo := 11; 									(* Set error number *)
			sErrorMsg := 'Synchronization plus reached';
		END_IF
	ELSE
		IF bSyncMinus
		THEN
			udnErrorNo := 12; 									(* Set error number *)
			sErrorMsg := 'Synchronization minus err';
		ELSIF bSyncPlus
		THEN
			udnErrorNo := 13; 									(* Set error number *)
			sErrorMsg := 'Synchronization plus err';
		END_IF
	END_IF

	bMoveToPlus := FALSE;			(* Move to plus direction *)
  	bMoveToMinus := FALSE;			(* Move to minus direction *)
	bTargetPlus := FALSE;
	bTargetMinus := FALSE;

END_IF

(* Check condition *)
tonConWatchDog(IN := (bMoveToMinus AND NOT bAtMinusLimit AND bAtPlusLimit)
					OR (bMoveToPlus AND bAtMinusLimit AND NOT bAtPlusLimit),
				PT := tConTimeOut);

IF tonConWatchDog.Q
    AND NOT bError
THEN
	IF bMoveToMinus
	    AND NOT bAtMinusLimit
	    AND bAtPlusLimit
	THEN
		udnErrorNo := 16; 									(* Set error number *)
		sErrorMsg := 'Direction minus not free.';

	ELSIF bMoveToPlus
		    AND bAtMinusLimit
		    AND NOT bAtPlusLimit
	THEN
		udnErrorNo := 17; 									(* Set error number *)
		sErrorMsg := 'Direction plus not free.';
	END_IF

	bMoveToPlus := FALSE;
	bMoveToMinus := FALSE;
	bTargetPlus := FALSE;
	bTargetMinus := FALSE;

END_IF

IF bExtAlarm
THEN
	udnErrorNo := 20; 									(* Set error number *)
	sErrorMsg := 'External alarm.';
END_IF

bError := udnErrorNo <> 0;


(* End plus position reached  *)
bLimitPlus := bAtPlusLimit
		       AND NOT bAtMinusLimit
		       AND NOT bError;

(* End minus position reached  *)
bLimitMinus := NOT bAtPlusLimit
		          AND bAtMinusLimit
		          AND NOT bError;

(* Motor off if error *)
IF bError
     AND (bMoveToPlus OR bMoveToMinus)
     AND bMotorCtrlErrOff
THEN
	bMoveToPlus := FALSE;			(* Move to plus direction *)
  	bMoveToMinus := FALSE;			(* Move to minus direction *)
	bTargetPlus := FALSE;
	bTargetMinus := FALSE;
END_IF

(* Check control off *)
IF bControlOff
   AND tControlOff > t#0ms
THEN
	tonControlOff(
		IN := bMoveToPlus OR bMoveToMinus
			OR bTargetPlus OR bTargetMinus,
		PT := tControlOff
	);

	IF tonControlOff.Q
	THEN
		bMoveToPlus := FALSE;
		bMoveToMinus := FALSE;
		bTargetPlus := FALSE;
		bTargetMinus := FALSE;
	END_IF;
    
ELSE
	tonControlOff(IN := FALSE);

	IF bControlOff
	    AND (
			bMoveToPlus OR bMoveToMinus
			OR bTargetPlus OR bTargetMinus
		      )
	THEN
		bMoveToPlus := FALSE;
		bMoveToMinus := FALSE;
		bTargetPlus := FALSE;
		bTargetMinus := FALSE;
	END_IF;
END_IF;

END_FUNCTION_BLOCK

// ---- POUs/Machine/Group_0500 - Transport/Gr05Control/Gr05Alarm/FB_Gr05Alarm.TcPOU
FUNCTION_BLOCK FB_Gr05Alarm
(*

The function block used to control general alarms of machine.

Constructor: 		Patryk Panylo
Company:		E. Riexinger GmbH
Date:			28.04.2015
Version:			1.00

Date:			Revision:		Who:				Comment
dd.mm.yyyy		x.xx			Initials			comment

*)
VAR_INPUT
	(* Input variables / Eingang Variablen *)
	etMachineMode				:ET_MachineMode;			(* Machine mode *)
	etMachineState				:ET_MachineState;			(* Machine state *)
	bNoEStop					:BOOL;						(* Emergency stop *)
	bConfirmAlarm				:BOOL;						(* Confirm alarm *)
	dtDateTime 					:DATE_AND_TIME;			(* Actual date and time *)
	nFatalErrorMaxIdx				:INT;						(* Maximal index of  using alarms *)
	nErrorMaxIdx					:INT;						(* Maximal index of  using alarms *)
	nWarningMaxIdx				:INT;						(* Maximal index of  using alarms *)
	nMessageMaxIdx				:INT;						(* Maximal index of  using alarms *)
	nHintMaxIdx					:INT;						(* Maximal index of  using alarms *)
	stAlarmIn						:ST_AlarmIn;					(* Alarm input *)
END_VAR
VAR_OUTPUT
	(* Output variables / Ausgang Variablen *)
	stAlarmOut					:ST_AlarmOut;				(* Alarm input *)
END_VAR
VAR_IN_OUT
	(* Input Output variables / Ausgang Variablen *)
	bMoveInterrupted				:BOOL;						(* Move interrupted *)
	bHomeCompleted				:BOOL;						(* Home completed *)
END_VAR
VAR
	(* Enummerations *)

	(* Variables *)

	(* References *)

	(* Interfaces *)

	(* Instances *)
	fbAlarm						:FB_Alarm;
END_VAR


(* Collection of alarms *)
fbAlarm(
	bEnable := TRUE,
	bNoEStop := bNoEStop,
	bReset := bConfirmAlarm,
	dtDateTime := dtDateTime,
	nFatalErrorMaxIdx := nFatalErrorMaxIdx,
	nErrorMaxIdx := nErrorMaxIdx,
	nWarningMaxIdx := nWarningMaxIdx,
	nMessageMaxIdx := nMessageMaxIdx,
	nHintMaxIdx := nHintMaxIdx,
    	stAlarmIn := stAlarmIn,
    	stAlarmOut => stAlarmOut
);

IF stAlarmOut.bFatalError
    OR stAlarmOut.bError
THEN
	(*bMoveInterrupted := FALSE;*)
	bHomeCompleted := FALSE;
END_IF;

END_FUNCTION_BLOCK

// ---- POUs/Machine/Group_0500 - Transport/Gr05Control/Gr05Safety/FB_Gr05Safety.TcPOU
FUNCTION_BLOCK FB_Gr05Safety
(*

The function block used to control genaeral safety of the machine.

Constructor: 		Patryk Panylo
Company:		E. Riexinger GmbH
Date:			28.04.2015
Version:			1.00

Date:			Revision:		Who:				Comment
dd.mm.yyyy		x.xx			Initials			comment

*)
VAR_INPUT
	(* Input variables / Eingang Variablen *)
	etMachineMode				:ET_MachineMode;			(* Machine mode *)
	etMachineState				:ET_MachineState;			(* Machine state *)
	bLightCurtain					:BOOL;						(* Light curtain ok / Freigabe Lichtschranke i.o *)
	bConfirmLightCurtain			:BOOL;						(* Confirm light Curtain input signal *)
	tLightCurtainDelay				:TIME := t#1s;					(* After time light Curtain safe *)
END_VAR
VAR_OUTPUT
	(* Output variables / Ausgang Variablen *)
	bLightCurtainOK				:BOOL;						(* Light curtain ok / Freigabe Lichtschranke i.o *)
	bConfirmedLightCurtain			:BOOL;						(* Confirmed light Curtain signal *)
	bNotInCrashArea				:BOOL;						(* Axis not in crash area with *)
END_VAR
VAR_IN_OUT
	(* Input Output variables / Ausgang Variablen *)

END_VAR
VAR
	(* Enummerations *)

	(* Variables *)

	(* References *)

	(* Interfaces *)

	(* Instances *)
	fbLightCurtain					:FB_LightCurtain;

END_VAR


A_LightCurtain();
A_SafetyArea();

ACTION A_LightCurtain:

(* Light Curtain control *)
fbLightCurtain(
	bEnable := TRUE,
	bIn := bLightCurtain,
	bInConf := bConfirmLightCurtain,
	tTimeOut := tLightCurtainDelay,
	bOut => bLightCurtainOK,
	bOutConf => bConfirmedLightCurtain
);
END_ACTION

ACTION A_SafetyArea:

(* Safety area *)
bNotInCrashArea := FALSE;

IF FALSE
THEN
	bNotInCrashArea := TRUE;
END_IF;
END_ACTION

END_FUNCTION_BLOCK

// ---- POUs/Machine/Group_0500 - Transport/Gr05Control/Gr05Signals/FB_Gr05Signals.TcPOU
FUNCTION_BLOCK FB_Gr05Signals
(*

The function block used to control general signals of the machine.

Constructor: 		Patryk Panylo
Company:		E. Riexinger GmbH
Date:			28.04.2015
Version:			1.00

Date:			Revision:		Who:				Comment
dd.mm.yyyy		x.xx			Initials			comment

*)
VAR_INPUT
	(* Input variables / Eingang Variablen *)
	etMachineMode				:ET_MachineMode;			(* Machine mode *)
	etMachineState				:ET_MachineState;			(* Machine state *)
	bMachineRunning				:BOOL;						(* Machine running / Maschine lauft *)
	bExecutedProcess			:BOOL;						(* Process executed *)
	stBlinker						:ST_Blinker;
END_VAR
VAR_OUTPUT
	(* Output variables / Ausgang Variablen *)
	bBulbBtnStop					:BOOL;						(* Signal button bulb "stop" / Signallampe "Stop" *)
	bBulbBtnStart					:BOOL;						(* Signal button bulb "start" / Signallampe "Start" *)
END_VAR
VAR_IN_OUT
	(* Input Output variables / Ausgang Variablen *)

END_VAR
VAR
	(* Enummerations *)

	(* Variables *)

	(* References *)

	(* Interfaces *)

	(* Instances *)
	fbSpindleHeadPresent			:FB_SignalHandlingDelay;
	fbFurrowingHeadPresent		:FB_SignalHandlingDelay;
END_VAR


A_SignalButton();

(*boutGr05PipeBeginEdge := binGr05PipeBeginEdge;*)

ACTION A_SignalButton:

(* Signal button bulb "stop" / Signallampe "Stop" *)
bBulbBtnStop := NOT bExecutedProcess;


(* Signal button bulb "start" / Signallampe "Start" *)
bBulbBtnStart := SEL(bExecutedProcess,
                           		     bMachineRunning AND stBlinker.Q1,
                           		     bMachineRunning);
END_ACTION

END_FUNCTION_BLOCK

// ---- POUs/Machine/Group_0500 - Transport/Gr05Control/Gr05Utility/FB_Gr05Utility.TcPOU
FUNCTION_BLOCK FB_Gr05Utility
(*

The function block used to control general utility of the machine.

Constructor: 		Patryk Panylo
Company:		E. Riexinger GmbH
Date:			28.04.2015
Version:			1.00

Date:			Revision:		Who:				Comment
dd.mm.yyyy		x.xx			Initials			comment

*)
VAR_INPUT
	(* Input variables / Eingang Variablen *)
	etMachineMode				:ET_MachineMode;			(* Machine mode *)
	etMachineState				:ET_MachineState;			(* Machine state *)
	bStartProcess				:BOOL;						(* Start process *)
	bStopProcess				:BOOL;						(* Stop process *)
	bSteppingProcess			:BOOL;						(* Stepping process *)
	bAutoCompleted				:BOOL;						(* Process completed *)
	bExeCounter					:BOOL;						(* Execute counter *)
	bStartTime					:BOOL;						(* Start measurement of cylce time *)
	bStopTime					:BOOL;						(* Stop measurement of cylce time *)
	bLifetimeOn					:BOOL;						(* Lifetime on *)
	bResetLifetimeAll				:BOOL; 						(* Reset all counters *)
	bResetLifetime				:BOOL;						(* Reset counter *)
	sLifetimeFilePath				:STRING;					(* File path for life time *)
	sLifetimeFileName			:STRING;					(* File name for life time *)
	bPipeEndEdgeIdentify			:BOOL;						(* Pipe end edge identify *)
	bPipeBeginEdgeIdentify		:BOOL;						(* Pipe begin edge identify *)
	rGlobalOverride				:REAL;						(* Global override *)
	tAdsTimeOut 					:TIME := t#2s;					(* Timout for ads commands *)
END_VAR
VAR_OUTPUT
	(* Output variables / Ausgang Variablen *)
	bExeProcess					:BOOL;						(* Execute process *)
	rActOverride					:REAL;						(* Actual override *)
	lrLifetimeAll					:LREAL;						(* Lifetime all *)
	lrLifetimeAfterReset			:LREAL;						(* Lifetime after reset *)
	lrLifetimeAfterTrunOn			:LREAL;						(* Lifetime after turn on *)
	bPipeEndPresent				:BOOL;						(* End of pipe present *)
	bPipeBeginPresent			:BOOL;						(* Begin of pipe present *)
END_VAR
VAR_IN_OUT
	(* Input Output variables / Ausgang Variablen *)
	bHomeCompleted				:BOOL;						(* Execute process *)
	rLocalOverride				:REAL;						(* Actual override *)
	udnCounterTotal				:UDINT;						(* Counter *)
END_VAR
VAR
	(* Enummerations *)

	(* Variables *)
	arudnCounterTotal				:ARRAY[0..1] OF UDINT;			(* Counter *)

	(* References *)

	(* Interfaces *)

	(* Instances *)
	fbStartProcess				:FB_StartProcess;
	fbOverride					:FB_Override;
	fbOverrideSelection			:FB_OverrideSelection;
	fbLifetime					:FB_TimeHoursCounter;		(* Machine lifetime *)
	arfbCounter					:ARRAY[0..1] OF FB_Counter;
	arfbCylceTime				:ARRAY[0..1] OF FB_Timer;
	fbPipeBeginIdentify			:FB_SignalHandlingEdge;
	fbPipeEndIdentify				:FB_SignalHandlingEdge;
END_VAR


A_StartProcess();
A_Override();
A_Counter();
A_CycleTime();
A_PipeIdentify();

ACTION A_Counter:

(* Hours counter *)
fbLifetime(
	bEnable := TRUE,
	bDeleteAll := bResetLifetimeAll,
	sAmsNetId := sgAmsNetId,
	bCount := bLifetimeOn,
	bSave := FALSE,
	bReset := bResetLifetime,
	sFilePath := sLifetimeFilePath,
	sFileName := sLifetimeFileName,
	tSaveIntervall := t#8m,
	tTimeout := tAdsTimeOut,
	lrAllOverHours => lrLifetimeAll,
	lrAfterResetHours => lrLifetimeAfterReset,
	lrNoRetainHours => lrLifetimeAfterTrunOn,
 );

(* Counter *)
arfbCounter[0](
	bEnable := TRUE,
	bExecute := bExeCounter,
	bReset := arfbCounter[0].bOverflow,
	udnCounter := udnCounterTotal
);

arfbCounter[1](
	bEnable := TRUE,
	bExecute := bExeCounter,
	bReset := arfbCounter[1].bOverflow,
	udnCounter := arudnCounterTotal[1]
);
END_ACTION

ACTION A_CycleTime:

(* Cylce time *)
arfbCylceTime[0](
	bEnable := TRUE,
	bReset := FALSE,
	bStartStop := bStartTime
			        AND bgGr00ModeAutomatic,
	bStop := bStopTime
		        OR bgGr00MachineStandstill,
	tMaxTime := t#480m,
	stRefTime => ,
	stActTime => ,
	stRestTime =>
);

arfbCylceTime[1](
	bEnable := TRUE,
	bReset := FALSE,
	bStartStop := bStartTime
			        AND bgGr00ModeAutomatic,
	bStop := bStopTime
		        OR bgGr00MachineStandstill,
	tMaxTime := t#480m,
	stRefTime => ,
	stActTime => ,
	stRestTime =>
);
END_ACTION

ACTION A_Override:

(* Override control *)
fbOverrideSelection(
	bEnable := TRUE,
	rGlobalOverride := rGlobalOverride,
	rLocalOverride := rLocalOverride
);

fbOverride(
	bEnable := TRUE,
	bBypassAccDec := etMachineMode = ET_MachineMode_eManual,
	rSetOverride := fbOverrideSelection.rActOverride,
	rAcc := rgGr05AdsOverrideAcc,
	rDec := rgGr00AdsOverrideDec,
	rActOverride => rActOverride
);
END_ACTION

ACTION A_PipeIdentify:

fbPipeEndIdentify(
	bEnable := TRUE,
	bIn := bPipeEndEdgeIdentify,
	tDelay := t#0s,
	bOut => bPipeEndPresent
);

fbPipeBeginIdentify(
	bEnable := TRUE,
	bIn := bPipeBeginEdgeIdentify,
	tDelay := t#0s,
	bOut => bPipeBeginPresent
);
END_ACTION

ACTION A_StartProcess:

(* Start auto process *)
fbStartProcess(
	bEnable := etMachineMode = ET_MachineMode_eAutomatic
			    OR etMachineMode = ET_MachineMode_eCycle
			    OR etMachineMode = ET_MachineMode_eStepping,
	bStart := bStartProcess,
	bStop := bStopProcess,
	bDone := bAutoCompleted,
	bStepping := bSteppingProcess,
	bHomeCompleted := bHomeCompleted,
	bStartProcess => bExeProcess
);
END_ACTION

END_FUNCTION_BLOCK

// ---- POUs/Machine/Group_0500 - Transport/Gr05HMI/Gr05HMI.TcPOU
PROGRAM Gr05HMI
VAR_INPUT
	(* Input variables / Eingang Variablen *)
	bEnable					:BOOL;						(* Enable Gr05HMI *)
END_VAR
VAR
	(* Enummerations *)

	(* Variables *)
	rOverride							:REAL;						(* Override 0 - 100 % *)
	lrManualVelo							:LREAL;						(* Manual velocity *)
	lrHomeVelo							:LREAL;						(* Home velocity *)
	lrAutoVelo							:LREAL;						(* Auto velocity *)
	udnCounterTotal						:UDINT;						(* Total counter *)

	lrOriginShiftPosAxisHE					:LREAL;											(* Origin shift position axis heating element [mm] *)
	lrHomePosAxisHE					:LREAL;											(* Home position axis heating element [mm] *)
	lrAxisHESoftLimitMax					:LREAL;											(* Software limit maximum axis heating element [mm] *)
	lrAxisHESoftLimitMin					:LREAL;											(* Software limit minimum axis heating element [mm] *)
	arunIRHSSetpoint						:ARRAY[1..nZONES_MAX_NO] OF LREAL;			(* IRHS setpoint *)
	arunPreHeatTime						:ARRAY[0..3] OF UINT;								(* PreHeat time [s] *)
	arunPreHeatPower					:ARRAY[0..3] OF UINT;								(* PreHeat power [%] *)
	arlrPreHeatTemp						:ARRAY[0..3] OF LREAL;							(* PreHeat temperatur [°] *)
	lrAxisHEPreHeatPos					:LREAL;											(* Heating element pre position [mm] *)
	lrShuttleBackForthDistance				:LREAL;											(* Shuttle distance between heating elemnt back and forth [mm] *)

	(* References *)

	(* Interfaces *)

	(* Instances *)

END_VAR

IF NOT bEnable
THEN
	RETURN;
END_IF;

A_GetHMIVar();
A_SetHMIVar();

ACTION A_GetHMIVar:

(* Collect hmi signals *)
;
END_ACTION

ACTION A_SetHMIVar:

